// TIA Portal project "M2471_Etiqueteuse" (V18)

(* hardware
DEVICE "Station S7-1200_1"  S7-1200 Station
   slot 0: "Châssis_0"  S7-1200 Rack  Rack  V1.0
   slot 1: "PLC_1"  CPU 1212C DC/DC/DC  6ES7 212-1AE40-0XB0  V4.5
   slot 2: "DI 16/DQ 16x24VDC_1"  6ES7 223-1BL32-0XB0  V2.0
DEVICE "HMI_1"  KTP700 Basic PN
   slot 0: "HMI_1"  KTP700 Basic PN  6AV2 123-2GB03-0AX0  13.0.1.0
   slot 1: "HMI_RT_2"  KTP700 Basic PN  6AV2 123-2GB03-0AX0  13.0.1.0
   slot 5: "HMI_1.IE_CP_1"  PROFINET Interface  13.0.1.0
      slot 1: "Interface PROFINET_1"  PROFINET Interface
         slot 1: "Port_1"  Port
*)

// ===== PLC "PLC_1"  CPU 1212C DC/DC/DC =====

VAR_GLOBAL   // PLC tag table "Table de variables standard"
   "Moteur_Con_Entree" AT %Q8.0 : Bool;
   "Moteur_Con_Etiquetage" AT %Q8.1 : Bool;
   "Moteur_Con_Sortie" AT %Q8.2 : Bool;
   "Moteur_Etiquetage" AT %Q0.7 : Bool;
   "Capteur_Con_Entree" AT %I0.2 : Bool;
   "Capteur_Etiquette" AT %I0.7 : Bool;
   "Capteur_Verin_Tete_Max" AT %I0.4 : Bool;
   "Capteur_Verin_Tete_Min" AT %I0.5 : Bool;
   "Capteur_Verin_Etiquette_Max" AT %I8.0 : Bool;
   "Findecourse_Entree_Petit" AT %I1.6 : Bool;
   "Findecourse_Entree_Grand" AT %I1.7 : Bool;
   "Findecourse_Hauteur_Haut" AT %I0.6 : Bool;
   "Relai_Securite_Arret" AT %I0.0 : Bool;
   "Relai_Secu" AT %Q0.0 : Bool;
   "Moteurpasapas_Haut" AT %M0.0 : Bool;
   "Moteurpasapas_Bas" AT %M0.1 : Bool;
   "Motor_EN" AT %Q0.2 : Bool;
   "Motor_CLK" AT %Q0.4 : Bool;
   "Motor_DIR" AT %Q0.3 : Bool;
   "Entre_Detection_Pot" AT %M0.2 : Bool;
   "Sortie_Detection_Pot" AT %M0.6 : Bool;
   "Butee_Bas_Calibration" AT %I0.1 : Bool;
   "Petit_Pot" AT %M1.0 : Bool;
   "Grand_Pot" AT %M1.1 : Bool;
   "retour_Menu" AT %M0.5 : Bool;
   "System_Byte" AT %MB2 : Byte;
   "FirstScan" AT %M2.0 : Bool;
   "DiagStatusUpdate" AT %M2.1 : Bool;
   "AlwaysTRUE" AT %M2.2 : Bool;
   "AlwaysFALSE" AT %M2.3 : Bool;
   "Clock_Byte" AT %MB3 : Byte;
   "Clock_10Hz" AT %M3.0 : Bool;
   "Clock_5Hz" AT %M3.1 : Bool;
   "Clock_2.5Hz" AT %M3.2 : Bool;
   "Clock_2Hz" AT %M3.3 : Bool;
   "Clock_1.25Hz" AT %M3.4 : Bool;
   "Clock_1Hz" AT %M3.5 : Bool;
   "Clock_0.625Hz" AT %M3.6 : Bool;
   "Clock_0.5Hz" AT %M3.7 : Bool;
   "System_Byte(1)" AT %MB1 : Byte;
   "Moteur_Pwm" AT %Q0.1 : Bool;
   "Controle_Verin" AT %Q8.3 : Bool;
   "Dir_Moteur_15v" AT %Q0.5 : Bool;
   "Detection_Sortie_Bas" AT %M9.2 : Bool;
   "Verin_Etiquette" AT %Q8.4 : Bool;
   "Detection_Entree_Bas" AT %I9.0 : Bool;
   "Detection_Entree_Haut" AT %I9.1 : Bool;
   "Findecourse_Sortie" AT %I9.2 : Bool;
   "Capteur_Position_Pot" AT %I0.3 : Bool;
   "Tag_1" AT %QW1008 : Int;
   "calibration" AT %M1.3 : Bool;
   "stop bourage" AT %M4.0 : Bool;
END_VAR

DATA_BLOCK "Bloc_M2471Etiqueteuse"   // DB1
{ S7_Optimized_Access := 'TRUE' }
VERSION : 0.1
   VAR
      Status_McPower : Bool;
      Hauteur_Haut_Manuel : Bool;
      P_Trig_Reset : Bool;
      Commande_Moteur_Etiquette : Bool;
      Hauteur_Bas_Manuel : Bool;
      Calibrage_Fini : Bool;
      Relai_Securite_Etat : Bool;
      Coordonees_Positionement : Int;
      Moteur_Hauteur_Etiquetage : Bool;
      Moteurpasapas_Sens : Bool;
      Stop_Etat : Bool;
      Moteur_Con_En : Bool;
      Moteur_Con_Et : Bool;
      Moteur_Con_So : Bool;
      Capteur_Entre : Bool;
      capteur_etiquette : Bool;
      Moteur_Etiquette : Bool;
      Capteur_Sortie : Bool;
      Detection_Entre_Petit : Bool;
      Detection_Sortie : Bool;
      Detection_Entre_Grand : Bool;
      Calibration_Home : Bool;
      SR_Home : Bool;
      Ajustement_Hauteur_G_P : Bool;
      Position_Done : Bool;
      Hauteur_Haut_G_P : Bool;
      Hauteur_Bas_G_P : Bool;
      SR_Correction : Bool;
      SR_position : Bool;
      Retour_Menu : Bool;
      Reset : Bool;
      Petit_Pot : Bool;
      Grand_Pot : Bool;
      SR_Position_Done : Bool;
      SR_Correction_Deplacement : Bool;
      Crorrection_Done : Bool;
      Prev_Hauteur_Haut_G_P : Bool;
      Prev_Hauteur_Bas_G_P : Bool;
      Dispense_Etiquette : Bool;
      SR_Etiquette : Bool;
      Etiquetage : Bool;
      P_Trig_Etiquetage : Bool;
      Calibration_set : Bool;
      SR_Home_1 : Bool;
      Sr_etiquetage2 : Bool;
      N_trig_Etiquette : Bool;
      P_trig_Calibration : Bool;
      Reset_Ton_Etiquetage : Bool;
      Controle_Verin_Etiquette : Bool;
      SR_Controle_Verin_Etiquette : Bool;
      Ouverture_Verin_Etiquette : Bool;
      P_trig_Verin_Etiquette : Bool;
      Detection_Petit_Pot : Bool;
      Detection_Grand_Pot : Bool;
      TON_Reset_Controle_Petit : Bool;
      TON_Reset_Controle_Grand : Bool;
      SR_Controle_Petit : Bool;
      SR_Controle_Grand : Bool;
      Sr_Capteur_Pot : Bool;
      P_Trig_Con_Entree : Bool;
      Sr_Capteur_Pot_2 : Bool;
      Sr_Serage_Pot : Bool;
      NTrig_Serage_Pot : Bool;
      SR_CON_Etiquetage : Bool;
      Timer_Con_Etiquetage : Bool;
      Etiquetage_Fini : Bool;
      Verin_Fin : Bool;
      SR_Controle_Verin : Bool;
      SR_Sortie : Bool;
      fin : Bool;
      P_trig_Con_Eti : Bool;
      p_trig_entre : Bool;
      N_trig_etiquetage : Bool;
      controle_Pwm : Bool;
      Machine_Etat : Int;
      Vue_Demarage : Bool;
      Vue_Bourage : Bool;
      Vue_Menu : Bool;
      Vue_Grand : Bool;
      Vue_Petit : Bool;
      Vue_Manuel : Bool;
      Vue_Advance : Bool;
      Bourage : Bool;
      Mise_En_Marche : Bool;
      SR_calibration_Fini : Bool;
      calibrer : Bool;
      Programe : Bool;
      Coordone_Petit_Pot : Int := 100;
      Coordone_Grand_Pot : Int := 160;
      Coordone_Manuel_Pot : Int;
      Confirmation_GP : Bool;
      Confirmation_PP : Bool;
      Pot_Correct : Bool;
      Pot_Incorect : Bool;
      Retour_Demarage : Bool;
      N_Trig_Relai : Bool;
      P_Trig_Reset_calibration : Bool;
      reset_calibration : Bool;
      P_Trig_pot_incorect : Bool;
      SR_Etiquetage_FP : Bool;
      reset_incorect : Bool;
      reset_state : Bool;
      SR_reset : Bool;
      changement_etiquette : Bool;
      nombre_Pot : Int;
      nombre_reset : Bool;
      nombre_limite : Int;
      nombre_Fini : Bool;
      Nombre_sans_limite : Bool;
      p_trigAjustement : Bool;
      p_trig_petit_grand : Bool;
      coordonee_ajustement : Int;
      p_trig_coordone_engage : Bool;
      SR_coordone_engage : Bool;
      p_trig_position_done : Bool;
      p_trig_deplacement : Bool;
      mode_advance : Bool;
      moteur_Grand_advance : Bool;
      moteur_Petit_advance : Bool;
      valeur_Grand_Advance : Int;
      valeur_Petit_Advance : Int;
      coordonne_advance : Int;
      Moteur_advance : Bool;
      Advance_trigger : Bool;
      coordonne_advance_mem : Int;
      valeur_advance_sup_g : Bool;
      valeur_advance_sup_p : Bool;
      p_trig_advance : Bool;
      Manuel_Mode : Bool;
      Manuel_set : Bool;
      Valeur_Manuel : Int;
      Bouton_Manuel_5 : Bool;
      Bouton_Manuel_10 : Bool;
      Bouton_Manuel_25 : Bool;
      Commande_Manuel : Bool;
      Bourage_Done : Bool;
      P_trig_Bourage : Bool;
      bourage_Pneumatique : Bool;
      validation_securite_1 : Bool;
      validation_securite_2 : Bool;
      Verin_Etiquetage : Bool;
      Verin_Etiquette : Bool;
      SR_Bourage_Relai_Secu : Bool;
      Securite_Verin : Bool;
      Home_Reset : Bool;
      p_Trig_Home_Reset : Bool;
      busy_home_Reset : Bool;
      Advance_SR_ajustement : Bool;
      Enable_avdance_Grand : Bool;
      Enable_avdance_Petit : Bool;
      Advance_Etiquetage : Bool;
      SR_Advance : Bool;
      Verin_Etiquetage_advance : Bool;
      Etiquetage_advance : Bool;
      SR_Verin_etiquetage : Bool;
      Bourage_Verin : Bool;
      SR_advance_coordone_done : Bool;
      bourage_verin_etiquette : Bool;
      SR_Grand_Advance : Bool;
      P_trig_Grand_Advance : Bool;
      SR_Petit_Advance : Bool;
      P_trig_Petit_Advance : Bool;
      Grand_Check_Advance : Bool;
      Petit_Check_Advance : Bool;
      Advance_Stop_G : Bool;
      Advance_Stop_P : Bool;
      SR_Controle_P : Bool;
      SR_Controle_G : Bool;
      sr_tapis_eti_fini : Bool;
      reset_Etiquetage : Bool;
      SR_reset_Eti : Bool;
      SR_incorect_tapis_verin : Bool;
      incorect_Reset_P : Bool;
      incorect_Reset_G : Bool;
      sr_con_sortie : Bool;
      Busy_Positionnement : Bool;
      SR_Etiquetage_stop : Bool;
      reset_Absolut_Positionement : Bool;
      error_Positionement : Bool;
      Postionement_reset_error : Bool;
      move_absolut_Busy_Advance : Bool;
      p_trig_advance_Move : Bool;
      p_trig_adv_Etiqu : Bool;
      "SR_advance reset" : Bool;
      SR_Busy_advance_done : Bool;
      advance_check_taille : Int;
      advance_trigger_engage : Bool;
      Sortie_1_etiquette : Bool;
      p_trig_Sortie_1_etiquette : Bool;
      Sr_Advance_fini : Bool;
      advance_move_done : Bool;
      SR_Reset_reset : Bool;
      reset_done : Bool;
      advance_time : Bool;
      advance_time_check : Bool;
      Valeur_manuel_bouton : Bool;
      SR_Manuel_Check : Bool;
      Input_Manuel : Bool;
      P_Trig_Vue_Manuel : Bool;
      reset_Manuel_Check : Bool;
      p_trig_bouton_manuel : Bool;
      insert_Manuel_hauteur : Bool;
      valeur_manuel_check : Int;
      coordoonee_positionement_manuel : Int;
      Etiquetage_comande : Bool;
      reset_sortie_con : Bool;
      SR_reset_con_sortie : Bool;
      p_trig_vue_menu : Bool;
      nouvelle_valeur_manuel : Int;
      comptage_advance_p : Int;
      comptage_advance_g : Int;
      reset_count_p : Bool;
      reset_count_g : Bool;
      bourage_reset : Bool;
      Sr_reset_engage : Bool;
      reset_busy : Bool;
      reset_execute : Bool;
      Sr_reset_done : Bool;
      reset_restart : Bool;
      Home_2_reset : Bool;
      p_trig_home : Bool;
      p_trig_bourage_done : Bool;
      Bourage_Hauteur : Bool;
      p_trig_bourage_hauteur : Bool;
      error_Positionement_Home : Bool;
      error_Positionement_GP : Bool;
      error_Positionement_auto : Bool;
      Fonction_reset : Bool;
      Petit_mem : Bool;
      Grand_mem : Bool;
      checking_taille : Bool;
      automatique_mem : Bool;
      automatique_petit : Bool;
      automatique_grand : Bool;
      set_preset_grand : Bool;
      set_preset_petit : Bool;
   END_VAR
BEGIN
END_DATA_BLOCK

DATA_BLOCK "Initialisation_DB"   // DB2
{ S7_Optimized_Access := 'TRUE' }
VERSION : 0.1
// stored: InstanceOfName Initialisation
"Initialisation"
BEGIN
END_DATA_BLOCK

DATA_BLOCK "En_Marche_DB"   // DB4
{ S7_Optimized_Access := 'TRUE' }
VERSION : 0.1
// stored: InstanceOfName Commande
"Commande"
BEGIN
END_DATA_BLOCK

DATA_BLOCK "HMI_AREA_POINTER"   // DB25
{ S7_Optimized_Access := 'TRUE' }
VERSION : 0.1
   VAR
      tache_API : Array[0..3] of Word;
      NumScreen : Int := 8;
   END_VAR
BEGIN
   tache_API[0] := 51;
   tache_API[2] := 0;
   tache_API[3] := 0;
   // tache_API[1] : Number Screen to display
END_DATA_BLOCK

DATA_BLOCK "Etat_&_Securite_DB"   // DB26
{ S7_Optimized_Access := 'TRUE' }
VERSION : 0.1
// stored: InstanceOfName Etat_&_Securite
"Etat_&_Securite"
BEGIN
END_DATA_BLOCK

DATA_BLOCK "Verin_DB"   // DB28
{ S7_Optimized_Access := 'TRUE' }
VERSION : 0.1
// stored: InstanceOfName Verin
"Verin"
BEGIN
END_DATA_BLOCK

DATA_BLOCK "Moteur_DB"   // DB30
{ S7_Optimized_Access := 'TRUE' }
VERSION : 0.1
// stored: InstanceOfName Moteur
"Moteur"
BEGIN
END_DATA_BLOCK

DATA_BLOCK "Controle_Etiquetage_DB"   // DB31
{ S7_Optimized_Access := 'TRUE' }
VERSION : 0.1
// stored: InstanceOfName Controle_Etiquetage
"Controle_Etiquetage"
BEGIN
END_DATA_BLOCK

DATA_BLOCK "Moteur_DB_1"   // DB35
{ S7_Optimized_Access := 'TRUE' }
VERSION : 0.1
// stored: InstanceOfName Moteur
"Moteur"
BEGIN
END_DATA_BLOCK

DATA_BLOCK "Commande_DB"   // DB37
{ S7_Optimized_Access := 'TRUE' }
VERSION : 0.1
// stored: InstanceOfName Commande
"Commande"
BEGIN
END_DATA_BLOCK

DATA_BLOCK "Commande_DB_1"   // DB38
{ S7_Optimized_Access := 'TRUE' }
VERSION : 0.1
// stored: InstanceOfName Commande
"Commande"
BEGIN
END_DATA_BLOCK

// folder: System blocks/Program resources

DATA_BLOCK "IEC_Timer_0_DB"   // DB5
{ S7_Optimized_Access := 'TRUE' }
AUTHOR : Simatic
FAMILY : IEC
NAME : IEC_TMR
VERSION : 1.0
// stored: InstanceOfName IEC_TIMER
"IEC_TIMER"
BEGIN
END_DATA_BLOCK

DATA_BLOCK "IEC_Counter_0_DB_1"   // DB6
{ S7_Optimized_Access := 'TRUE' }
AUTHOR : Simatic
FAMILY : IEC
NAME : CNTR
VERSION : 1.0
// stored: InstanceOfName IEC_COUNTER
"IEC_COUNTER"
BEGIN
END_DATA_BLOCK

DATA_BLOCK "IEC_Timer_0_DB_2"   // DB7
{ S7_Optimized_Access := 'TRUE' }
AUTHOR : Simatic
FAMILY : IEC
NAME : IEC_TMR
VERSION : 1.0
// stored: InstanceOfName IEC_TIMER
"IEC_TIMER"
BEGIN
END_DATA_BLOCK

DATA_BLOCK "IEC_Timer_0_DB_3"   // DB10
{ S7_Optimized_Access := 'TRUE' }
AUTHOR : Simatic
FAMILY : IEC
NAME : IEC_TMR
VERSION : 1.0
// stored: InstanceOfName IEC_TIMER
"IEC_TIMER"
BEGIN
END_DATA_BLOCK

DATA_BLOCK "IEC_Timer_0_DB_4"   // DB13
{ S7_Optimized_Access := 'TRUE' }
AUTHOR : Simatic
FAMILY : IEC
NAME : IEC_TMR
VERSION : 1.0
// stored: InstanceOfName IEC_TIMER
"IEC_TIMER"
BEGIN
END_DATA_BLOCK

DATA_BLOCK "IEC_Timer_0_DB_5"   // DB15
{ S7_Optimized_Access := 'TRUE' }
AUTHOR : Simatic
FAMILY : IEC
NAME : IEC_TMR
VERSION : 1.0
// stored: InstanceOfName IEC_TIMER
"IEC_TIMER"
BEGIN
END_DATA_BLOCK

DATA_BLOCK "IEC_Counter_0_DB_2"   // DB16
{ S7_Optimized_Access := 'TRUE' }
AUTHOR : Simatic
FAMILY : IEC
NAME : CNTR
VERSION : 1.0
// stored: InstanceOfName IEC_COUNTER
"IEC_COUNTER"
BEGIN
END_DATA_BLOCK

DATA_BLOCK "IEC_Timer_0_DB_7"   // DB17
{ S7_Optimized_Access := 'TRUE' }
AUTHOR : Simatic
FAMILY : IEC
NAME : IEC_TMR
VERSION : 1.0
// stored: InstanceOfName IEC_TIMER
"IEC_TIMER"
BEGIN
END_DATA_BLOCK

DATA_BLOCK "IEC_Timer_0_DB_8"   // DB18
{ S7_Optimized_Access := 'TRUE' }
AUTHOR : Simatic
FAMILY : IEC
NAME : IEC_TMR
VERSION : 1.0
// stored: InstanceOfName IEC_TIMER
"IEC_TIMER"
BEGIN
END_DATA_BLOCK

DATA_BLOCK "IEC_Counter_0_DB"   // DB20
{ S7_Optimized_Access := 'TRUE' }
AUTHOR : Simatic
FAMILY : IEC
NAME : CNTR
VERSION : 1.0
// stored: InstanceOfName IEC_COUNTER
"IEC_COUNTER"
BEGIN
END_DATA_BLOCK

DATA_BLOCK "IEC_Timer_0_DB_9"   // DB27
{ S7_Optimized_Access := 'TRUE' }
AUTHOR : Simatic
FAMILY : IEC
NAME : IEC_TMR
VERSION : 1.0
// stored: InstanceOfName IEC_TIMER
"IEC_TIMER"
BEGIN
END_DATA_BLOCK

DATA_BLOCK "IEC_Timer_0_DB_10"   // DB29
{ S7_Optimized_Access := 'TRUE' }
AUTHOR : Simatic
FAMILY : IEC
NAME : IEC_TMR
VERSION : 1.0
// stored: InstanceOfName IEC_TIMER
"IEC_TIMER"
BEGIN
END_DATA_BLOCK

DATA_BLOCK "IEC_Timer_0_DB_11"   // DB32
{ S7_Optimized_Access := 'TRUE' }
AUTHOR : Simatic
FAMILY : IEC
NAME : IEC_TMR
VERSION : 1.0
// stored: InstanceOfName IEC_TIMER
"IEC_TIMER"
BEGIN
END_DATA_BLOCK

DATA_BLOCK "IEC_Timer_0_DB_12"   // DB34
{ S7_Optimized_Access := 'TRUE' }
AUTHOR : Simatic
FAMILY : IEC
NAME : IEC_TMR
VERSION : 1.0
// stored: InstanceOfName IEC_TIMER
"IEC_TIMER"
BEGIN
END_DATA_BLOCK

DATA_BLOCK "IEC_Timer_0_DB_14"   // DB36
{ S7_Optimized_Access := 'TRUE' }
AUTHOR : Simatic
FAMILY : IEC
NAME : IEC_TMR
VERSION : 1.0
// stored: InstanceOfName IEC_TIMER
"IEC_TIMER"
BEGIN
END_DATA_BLOCK

DATA_BLOCK "IEC_Timer_0_DB_17"   // DB39
{ S7_Optimized_Access := 'TRUE' }
AUTHOR : Simatic
FAMILY : IEC
NAME : IEC_TMR
VERSION : 1.0
// stored: InstanceOfName IEC_TIMER
"IEC_TIMER"
BEGIN
END_DATA_BLOCK

DATA_BLOCK "IEC_Timer_0_DB_18"   // DB40
{ S7_Optimized_Access := 'TRUE' }
AUTHOR : Simatic
FAMILY : IEC
NAME : IEC_TMR
VERSION : 1.0
// stored: InstanceOfName IEC_TIMER
"IEC_TIMER"
BEGIN
END_DATA_BLOCK

DATA_BLOCK "IEC_Timer_0_DB_19"   // DB41
{ S7_Optimized_Access := 'TRUE' }
AUTHOR : Simatic
FAMILY : IEC
NAME : IEC_TMR
VERSION : 1.0
// stored: InstanceOfName IEC_TIMER
"IEC_TIMER"
BEGIN
END_DATA_BLOCK

DATA_BLOCK "IEC_Timer_0_DB_20"   // DB42
{ S7_Optimized_Access := 'TRUE' }
AUTHOR : Simatic
FAMILY : IEC
NAME : IEC_TMR
VERSION : 1.0
// stored: InstanceOfName IEC_TIMER
"IEC_TIMER"
BEGIN
END_DATA_BLOCK

DATA_BLOCK "IEC_Timer_0_DB_21"   // DB45
{ S7_Optimized_Access := 'TRUE' }
AUTHOR : Simatic
FAMILY : IEC
NAME : IEC_TMR
VERSION : 1.0
// stored: InstanceOfName IEC_TIMER
"IEC_TIMER"
BEGIN
END_DATA_BLOCK

DATA_BLOCK "IEC_Timer_0_DB_22"   // DB46
{ S7_Optimized_Access := 'TRUE' }
AUTHOR : Simatic
FAMILY : IEC
NAME : IEC_TMR
VERSION : 1.0
// stored: InstanceOfName IEC_TIMER
"IEC_TIMER"
BEGIN
END_DATA_BLOCK

DATA_BLOCK "IEC_Timer_0_DB_23"   // DB47
{ S7_Optimized_Access := 'TRUE' }
AUTHOR : Simatic
FAMILY : IEC
NAME : IEC_TMR
VERSION : 1.0
// stored: InstanceOfName IEC_TIMER
"IEC_TIMER"
BEGIN
END_DATA_BLOCK

DATA_BLOCK "IEC_Timer_0_DB_24"   // DB48
{ S7_Optimized_Access := 'TRUE' }
AUTHOR : Simatic
FAMILY : IEC
NAME : IEC_TMR
VERSION : 1.0
// stored: InstanceOfName IEC_TIMER
"IEC_TIMER"
BEGIN
END_DATA_BLOCK

// folder: (top level)

DATA_BLOCK "Axe_1"   // DB8, Motion_DB
{ S7_Optimized_Access := 'TRUE' }
AUTHOR : SIMATIC
FAMILY : BasicMC
NAME : TO_PosAx
VERSION : 8.0
// stored: InstanceOfName TO_PositioningAxis
"TO_PositioningAxis"
BEGIN
   // Axis.PositionLimitsMin_AddressCU = %I0.1
   // Axis.PositionLimitsMax_AddressCU = %I0.6
   // Axis.DirectionOutputEnabledCU = TRUE
   // Axis.LengthUnitNormalized.Distance = 1013
   // Axis.HomingReferencePointSwitch_AddressCU = %I0.1
   // Axis.EnableOutput_AddressCU = %Q0.2
   // Axis.OnlinePtoModeCU = 16#0000_0002
   // Axis.SelectedChannel2EnumCU = %Q0.3
   // Axis.SelectedChannel1EnumCU = %Q0.4
   // Pulse.MinDeltaDeltaFrequencyCU = 0.004
   // Pulse.MaxDeltaDeltaFrequencyCU = 1.0E+10
   // Pulse.MinDeltaFrequencyCU = 0.005
   // Pulse.MaxDeltaFrequencyCU = 9.5E+9
   // Pulse.MinFrequencyCU = 1.0
   // Pulse.MaxFrequencyCU = 30000.0
   // Pulse.OutputSourceCU = 16#0000_0000
   // Axis.SelectPTO = 0
END_DATA_BLOCK

FUNCTION_BLOCK "Etat_&_Securite"   // FB1, LAD
{ S7_Optimized_Access := 'TRUE' }
VERSION : 0.1
   VAR_TEMP   // added for the SCL form of the ladder/FBD networks
      _w1 : Bool;
      _w2 : Bool;
   END_VAR
BEGIN

REGION Network 1: Relai de Secrurite
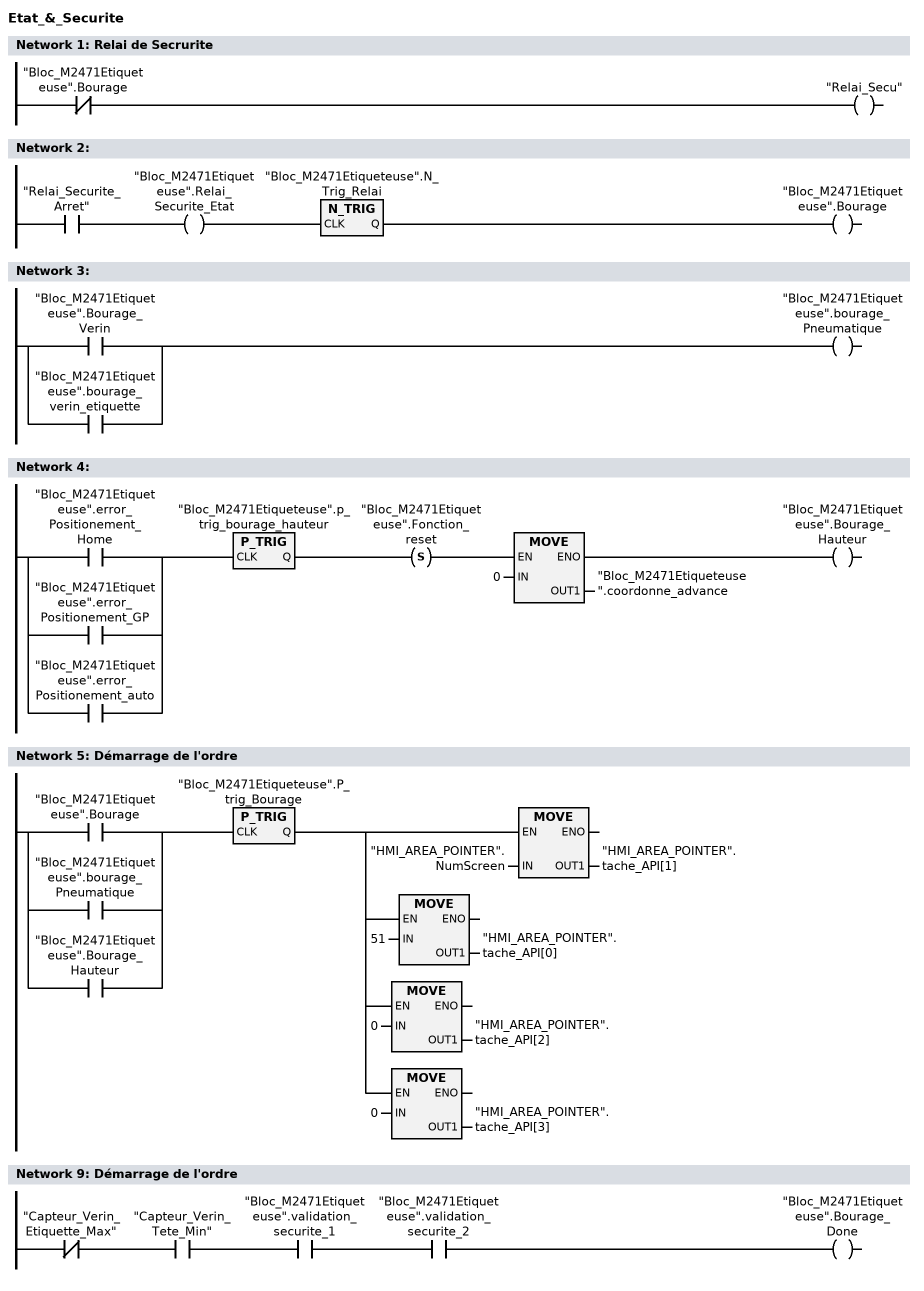
   RUNG wire#powerrail
      I_Contact( "Bloc_M2471Etiqueteuse".Bourage )
      Coil( "Relai_Secu" )
   END_RUNG
   // the same network as SCL:
   "Relai_Secu" := NOT "Bloc_M2471Etiqueteuse".Bourage;
END_REGION

REGION Network 2
   RUNG wire#powerrail
      Contact( "Relai_Securite_Arret" )
      Coil( "Bloc_M2471Etiqueteuse".Relai_Securite_Etat )
      N_Trig( "Bloc_M2471Etiqueteuse".N_Trig_Relai )
      Coil( "Bloc_M2471Etiqueteuse".Bourage )
   END_RUNG
   // the same network as SCL:
   "Bloc_M2471Etiqueteuse".Relai_Securite_Etat := "Relai_Securite_Arret";
   #_w1 := NOT "Relai_Securite_Arret" AND "Bloc_M2471Etiqueteuse".N_Trig_Relai;   // falling edge
   "Bloc_M2471Etiqueteuse".N_Trig_Relai := "Relai_Securite_Arret";
   "Bloc_M2471Etiqueteuse".Bourage := #_w1;
END_REGION

REGION Network 3
   RUNG wire#powerrail
      Contact( "Bloc_M2471Etiqueteuse".Bourage_Verin )
      wire#w1
      Coil( "Bloc_M2471Etiqueteuse".bourage_Pneumatique )
   END_RUNG
   RUNG wire#powerrail
      Contact( "Bloc_M2471Etiqueteuse".bourage_verin_etiquette )
   END_RUNG wire#w1
   // the same network as SCL:
   "Bloc_M2471Etiqueteuse".bourage_Pneumatique := "Bloc_M2471Etiqueteuse".Bourage_Verin OR "Bloc_M2471Etiqueteuse".bourage_verin_etiquette;
END_REGION

REGION Network 4
   RUNG wire#powerrail
      Contact( "Bloc_M2471Etiqueteuse".error_Positionement_Home )
      wire#w1
      P_Trig( "Bloc_M2471Etiqueteuse".p_trig_bourage_hauteur )
      S_Coil( "Bloc_M2471Etiqueteuse".Fonction_reset )
      Move(in := 0, out1 => "Bloc_M2471Etiqueteuse".coordonne_advance)
      Coil( "Bloc_M2471Etiqueteuse".Bourage_Hauteur )
   END_RUNG
   RUNG wire#powerrail
      Contact( "Bloc_M2471Etiqueteuse".error_Positionement_GP )
   END_RUNG wire#w1
   RUNG wire#powerrail
      Contact( "Bloc_M2471Etiqueteuse".error_Positionement_auto )
   END_RUNG wire#w1
   // the same network as SCL:
   #_w1 := "Bloc_M2471Etiqueteuse".error_Positionement_Home OR "Bloc_M2471Etiqueteuse".error_Positionement_GP OR "Bloc_M2471Etiqueteuse".error_Positionement_auto;
   #_w2 := #_w1 AND NOT "Bloc_M2471Etiqueteuse".p_trig_bourage_hauteur;   // rising edge
   "Bloc_M2471Etiqueteuse".p_trig_bourage_hauteur := #_w1;
   IF #_w2 THEN
       "Bloc_M2471Etiqueteuse".Fonction_reset := TRUE;
       "Bloc_M2471Etiqueteuse".coordonne_advance := 0;
   END_IF;
   "Bloc_M2471Etiqueteuse".Bourage_Hauteur := #_w2;
END_REGION

REGION Network 5: Démarrage de l'ordre
   RUNG wire#powerrail
      Contact( "Bloc_M2471Etiqueteuse".Bourage )
      wire#w1
      P_Trig( "Bloc_M2471Etiqueteuse".P_trig_Bourage )
      wire#w2
      Move(in := "HMI_AREA_POINTER".NumScreen, out1 => "HMI_AREA_POINTER".tache_API[1])
   END_RUNG
   RUNG wire#powerrail
      Contact( "Bloc_M2471Etiqueteuse".bourage_Pneumatique )
   END_RUNG wire#w1
   RUNG wire#powerrail
      Contact( "Bloc_M2471Etiqueteuse".Bourage_Hauteur )
   END_RUNG wire#w1
   RUNG wire#w2
      Move(in := 51, out1 => "HMI_AREA_POINTER".tache_API[0])
   END_RUNG
   RUNG wire#w2
      Move(in := 0, out1 => "HMI_AREA_POINTER".tache_API[2])
   END_RUNG
   RUNG wire#w2
      Move(in := 0, out1 => "HMI_AREA_POINTER".tache_API[3])
   END_RUNG
   // the same network as SCL:
   #_w1 := "Bloc_M2471Etiqueteuse".Bourage OR "Bloc_M2471Etiqueteuse".bourage_Pneumatique OR "Bloc_M2471Etiqueteuse".Bourage_Hauteur;
   #_w2 := #_w1 AND NOT "Bloc_M2471Etiqueteuse".P_trig_Bourage;   // rising edge
   "Bloc_M2471Etiqueteuse".P_trig_Bourage := #_w1;
   IF #_w2 THEN
       "HMI_AREA_POINTER".tache_API[1] := "HMI_AREA_POINTER".NumScreen;
       "HMI_AREA_POINTER".tache_API[0] := 51;
       "HMI_AREA_POINTER".tache_API[2] := 0;
       "HMI_AREA_POINTER".tache_API[3] := 0;
   END_IF;
END_REGION

REGION Network 6 (SCL): Machine Etat
   IF "Relai_Securite_Arret" = FALSE OR "Bloc_M2471Etiqueteuse".Bourage OR "Bloc_M2471Etiqueteuse".Bourage_Hauteur OR "Bloc_M2471Etiqueteuse".bourage_Pneumatique OR "Bloc_M2471Etiqueteuse".bourage_reset THEN
       "Bloc_M2471Etiqueteuse".Machine_Etat := 0;

   ELSIF "Bloc_M2471Etiqueteuse".Machine_Etat = 0 AND "Relai_Securite_Arret" = TRUE AND "Bloc_M2471Etiqueteuse".Relai_Securite_Etat = TRUE AND NOT "Bloc_M2471Etiqueteuse".Vue_Bourage =  TRUE THEN
       "Bloc_M2471Etiqueteuse".Machine_Etat := 1;

   ELSIF "Bloc_M2471Etiqueteuse".Machine_Etat = 1 AND "Bloc_M2471Etiqueteuse".calibrer = 1 THEN
      "Bloc_M2471Etiqueteuse".Machine_Etat := 2;

   ELSIF "Bloc_M2471Etiqueteuse".Machine_Etat = 2 AND "Bloc_M2471Etiqueteuse".Programe = 1 THEN
       "Bloc_M2471Etiqueteuse".Machine_Etat := 3;

   ELSIF "Bloc_M2471Etiqueteuse".Machine_Etat = 3 AND "Bloc_M2471Etiqueteuse".Programe = 0 THEN
       "Bloc_M2471Etiqueteuse".Machine_Etat := 2;
   END_IF;
END_REGION

REGION Network 7 (SCL): Etat et Variable
   IF "Bloc_M2471Etiqueteuse".Machine_Etat = 0 THEN
       "Bloc_M2471Etiqueteuse".Calibration_set := 0;
       "Bloc_M2471Etiqueteuse".reset_state := 0;
       "Bloc_M2471Etiqueteuse".Mise_En_Marche := FALSE;

   ELSIF "Bloc_M2471Etiqueteuse".Machine_Etat = 1 THEN
       "Bloc_M2471Etiqueteuse".Fonction_reset :=0;
       "Bloc_M2471Etiqueteuse".Calibration_set := 1;
       "Bloc_M2471Etiqueteuse".reset_state := 0;
       "Bloc_M2471Etiqueteuse".Mise_En_Marche := FALSE;

   ELSIF "Bloc_M2471Etiqueteuse".Machine_Etat = 2 THEN
       "Bloc_M2471Etiqueteuse".Calibration_set := 0;
       "Bloc_M2471Etiqueteuse".reset_state := 0;
       "Bloc_M2471Etiqueteuse".Mise_En_Marche := FALSE;

   ELSIF "Bloc_M2471Etiqueteuse".Machine_Etat = 3 THEN
       "Bloc_M2471Etiqueteuse".reset_state := 1;
       "Bloc_M2471Etiqueteuse".Mise_En_Marche := TRUE;

   END_IF;
END_REGION

REGION Network 8 (SCL): Programmes
   IF "Bloc_M2471Etiqueteuse".Vue_Bourage OR "Bloc_M2471Etiqueteuse".Vue_Demarage = 1 OR "Bloc_M2471Etiqueteuse".Vue_Menu = 1 THEN
       "Bloc_M2471Etiqueteuse".Programe := 0;

   ELSIF "Bloc_M2471Etiqueteuse".Vue_Grand = 1 OR "Bloc_M2471Etiqueteuse".Vue_Petit = 1 OR "Bloc_M2471Etiqueteuse".Vue_Manuel = 1 THEN
       "Bloc_M2471Etiqueteuse".Programe := 1;

   ELSIF "Bloc_M2471Etiqueteuse".Vue_Advance = 1 THEN
       "Bloc_M2471Etiqueteuse".Programe := 1;
       "Bloc_M2471Etiqueteuse".mode_advance := 1;

   END_IF;
END_REGION

REGION Network 9: Démarrage de l'ordre
   RUNG wire#powerrail
      I_Contact( "Capteur_Verin_Etiquette_Max" )
      Contact( "Capteur_Verin_Tete_Min" )
      Contact( "Bloc_M2471Etiqueteuse".validation_securite_1 )
      Contact( "Bloc_M2471Etiqueteuse".validation_securite_2 )
      Coil( "Bloc_M2471Etiqueteuse".Bourage_Done )
   END_RUNG
   // the same network as SCL:
   "Bloc_M2471Etiqueteuse".Bourage_Done := NOT "Capteur_Verin_Etiquette_Max" AND "Capteur_Verin_Tete_Min" AND "Bloc_M2471Etiqueteuse".validation_securite_1 AND "Bloc_M2471Etiqueteuse".validation_securite_2;
END_REGION
END_FUNCTION_BLOCK

FUNCTION_BLOCK "Verin"   // FB2, LAD
{ S7_Optimized_Access := 'TRUE' }
VERSION : 0.1
   VAR_TEMP   // added for the SCL form of the ladder/FBD networks
      _w1 : Bool;
      _w2 : Bool;
      _w3 : Bool;
   END_VAR
BEGIN

REGION Network 1
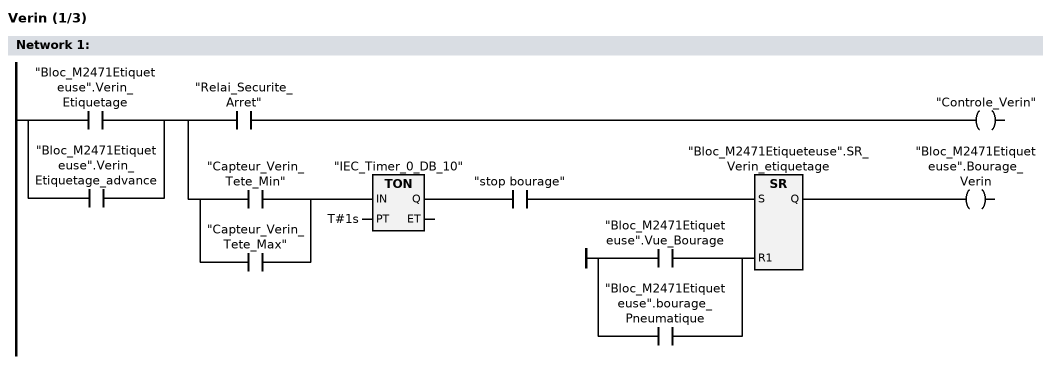
   #_w1 := "Bloc_M2471Etiqueteuse".Verin_Etiquetage OR "Bloc_M2471Etiqueteuse".Verin_Etiquetage_advance;
   "Controle_Verin" := #_w1 AND "Relai_Securite_Arret";
   "IEC_Timer_0_DB_10".TON(IN := #_w1 AND ("Capteur_Verin_Tete_Min" OR "Capteur_Verin_Tete_Max"), PT := T#1s);
   IF "IEC_Timer_0_DB_10".Q AND "stop bourage" THEN
       "Bloc_M2471Etiqueteuse".SR_Verin_etiquetage := TRUE;   // SR flip-flop
   END_IF;
   IF "Bloc_M2471Etiqueteuse".Vue_Bourage OR "Bloc_M2471Etiqueteuse".bourage_Pneumatique THEN
       "Bloc_M2471Etiqueteuse".SR_Verin_etiquetage := FALSE;
   END_IF;
   "Bloc_M2471Etiqueteuse".Bourage_Verin := "Bloc_M2471Etiqueteuse".SR_Verin_etiquetage;
END_REGION

REGION Network 2: commande Pneumatique Verin et tapsi etiquetage
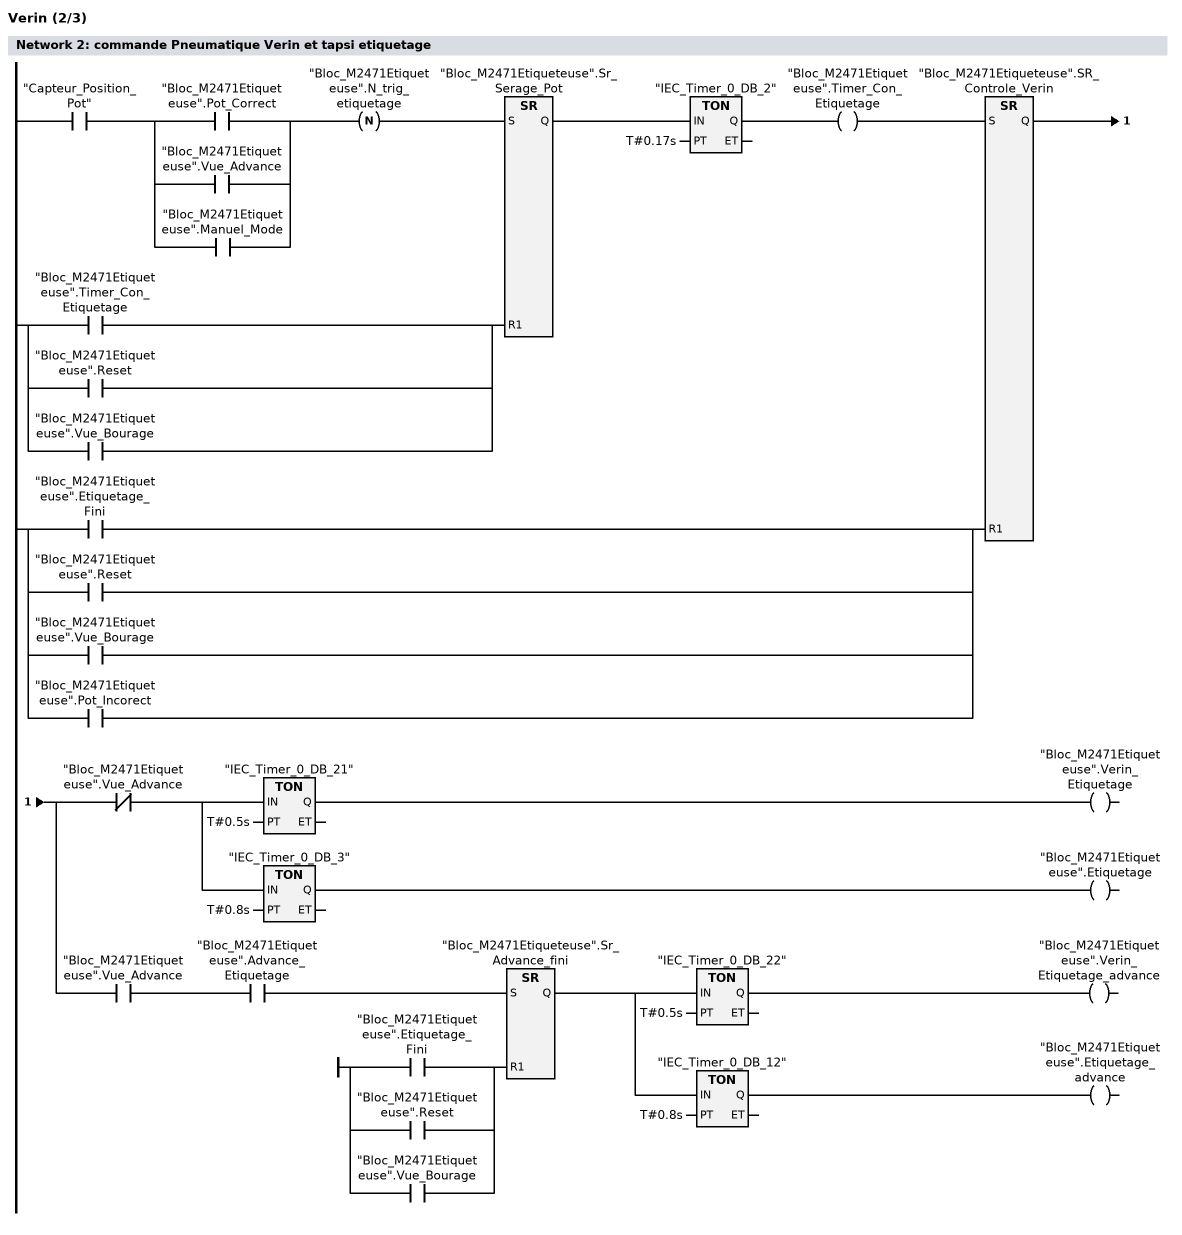
   #_w1 := "Capteur_Position_Pot" AND ("Bloc_M2471Etiqueteuse".Pot_Correct OR "Bloc_M2471Etiqueteuse".Vue_Advance OR "Bloc_M2471Etiqueteuse".Manuel_Mode);
   #_w2 := NOT #_w1 AND "Bloc_M2471Etiqueteuse".N_trig_etiquetage;   // falling edge
   "Bloc_M2471Etiqueteuse".N_trig_etiquetage := #_w1;
   IF #_w2 THEN
       "Bloc_M2471Etiqueteuse".Sr_Serage_Pot := TRUE;   // SR flip-flop
   END_IF;
   IF "Bloc_M2471Etiqueteuse".Timer_Con_Etiquetage OR "Bloc_M2471Etiqueteuse".Reset OR "Bloc_M2471Etiqueteuse".Vue_Bourage THEN
       "Bloc_M2471Etiqueteuse".Sr_Serage_Pot := FALSE;
   END_IF;
   "IEC_Timer_0_DB_2".TON(IN := "Bloc_M2471Etiqueteuse".Sr_Serage_Pot, PT := T#0.17s);
   "Bloc_M2471Etiqueteuse".Timer_Con_Etiquetage := "IEC_Timer_0_DB_2".Q;
   IF "IEC_Timer_0_DB_2".Q THEN
       "Bloc_M2471Etiqueteuse".SR_Controle_Verin := TRUE;   // SR flip-flop
   END_IF;
   IF "Bloc_M2471Etiqueteuse".Etiquetage_Fini OR "Bloc_M2471Etiqueteuse".Reset OR "Bloc_M2471Etiqueteuse".Vue_Bourage OR "Bloc_M2471Etiqueteuse".Pot_Incorect THEN
       "Bloc_M2471Etiqueteuse".SR_Controle_Verin := FALSE;
   END_IF;
   #_w3 := "Bloc_M2471Etiqueteuse".SR_Controle_Verin AND NOT "Bloc_M2471Etiqueteuse".Vue_Advance;
   "IEC_Timer_0_DB_21".TON(IN := #_w3, PT := T#0.5s);
   "Bloc_M2471Etiqueteuse".Verin_Etiquetage := "IEC_Timer_0_DB_21".Q;
   "IEC_Timer_0_DB_3".TON(IN := #_w3, PT := T#0.8s);
   "Bloc_M2471Etiqueteuse".Etiquetage := "IEC_Timer_0_DB_3".Q;
   IF "Bloc_M2471Etiqueteuse".SR_Controle_Verin AND "Bloc_M2471Etiqueteuse".Vue_Advance AND "Bloc_M2471Etiqueteuse".Advance_Etiquetage THEN
       "Bloc_M2471Etiqueteuse".Sr_Advance_fini := TRUE;   // SR flip-flop
   END_IF;
   IF "Bloc_M2471Etiqueteuse".Etiquetage_Fini OR "Bloc_M2471Etiqueteuse".Reset OR "Bloc_M2471Etiqueteuse".Vue_Bourage THEN
       "Bloc_M2471Etiqueteuse".Sr_Advance_fini := FALSE;
   END_IF;
   "IEC_Timer_0_DB_22".TON(IN := "Bloc_M2471Etiqueteuse".Sr_Advance_fini, PT := T#0.5s);
   "Bloc_M2471Etiqueteuse".Verin_Etiquetage_advance := "IEC_Timer_0_DB_22".Q;
   "IEC_Timer_0_DB_12".TON(IN := "Bloc_M2471Etiqueteuse".Sr_Advance_fini, PT := T#0.8s);
   "Bloc_M2471Etiqueteuse".Etiquetage_advance := "IEC_Timer_0_DB_12".Q;
END_REGION

REGION Network 3
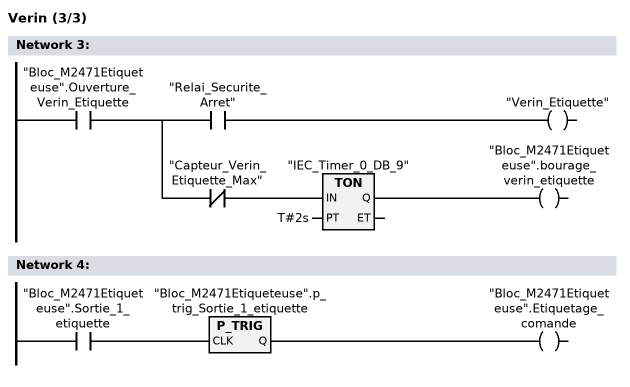
   "Verin_Etiquette" := "Bloc_M2471Etiqueteuse".Ouverture_Verin_Etiquette AND "Relai_Securite_Arret";
   "IEC_Timer_0_DB_9".TON(IN := "Bloc_M2471Etiqueteuse".Ouverture_Verin_Etiquette AND NOT "Capteur_Verin_Etiquette_Max",
                          PT := T#2s);
   "Bloc_M2471Etiqueteuse".bourage_verin_etiquette := "IEC_Timer_0_DB_9".Q;
END_REGION

REGION Network 4
   RUNG wire#powerrail
      Contact( "Bloc_M2471Etiqueteuse".Sortie_1_etiquette )
      P_Trig( "Bloc_M2471Etiqueteuse".p_trig_Sortie_1_etiquette )
      Coil( "Bloc_M2471Etiqueteuse".Etiquetage_comande )
   END_RUNG
   // the same network as SCL:
   #_w1 := "Bloc_M2471Etiqueteuse".Sortie_1_etiquette AND NOT "Bloc_M2471Etiqueteuse".p_trig_Sortie_1_etiquette;   // rising edge
   "Bloc_M2471Etiqueteuse".p_trig_Sortie_1_etiquette := "Bloc_M2471Etiqueteuse".Sortie_1_etiquette;
   "Bloc_M2471Etiqueteuse".Etiquetage_comande := #_w1;
END_REGION
END_FUNCTION_BLOCK

FUNCTION_BLOCK "Commande"   // FB3, LAD
{ S7_Optimized_Access := 'TRUE' }
VERSION : 0.1
   VAR_INPUT
      Valeur_Petit : Int;
      Valeur_Grand : Int;
      Valeur_Ajustement : Int;
   END_VAR
   VAR_TEMP   // added for the SCL form of the ladder/FBD networks
      _w1 : Bool;
   END_VAR
BEGIN

REGION Network 1: Reset
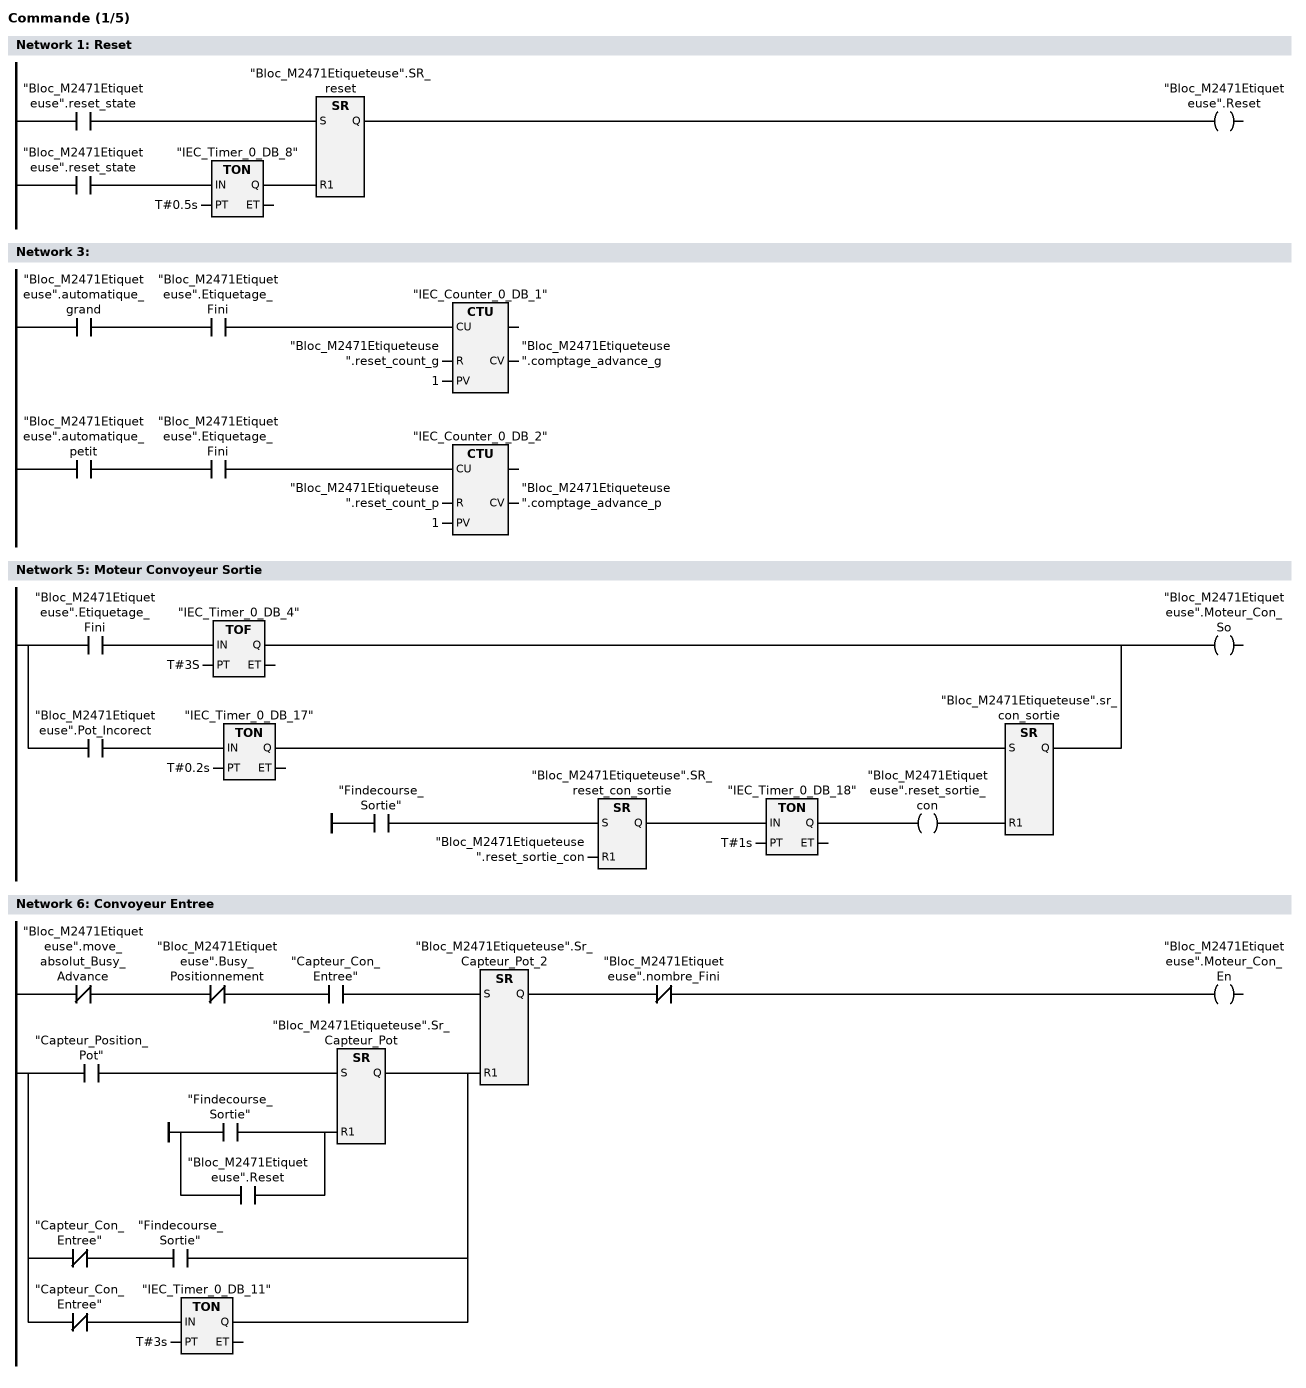
   "IEC_Timer_0_DB_8".TON(IN := "Bloc_M2471Etiqueteuse".reset_state, PT := T#0.5s);
   IF "Bloc_M2471Etiqueteuse".reset_state THEN
       "Bloc_M2471Etiqueteuse".SR_reset := TRUE;   // SR flip-flop
   END_IF;
   IF "IEC_Timer_0_DB_8".Q THEN "Bloc_M2471Etiqueteuse".SR_reset := FALSE; END_IF;
   "Bloc_M2471Etiqueteuse".Reset := "Bloc_M2471Etiqueteuse".SR_reset;
END_REGION

REGION Network 2 (SCL): detection grand ou petit pot ou automatique
   IF "Detection_Entree_Bas" OR "Detection_Entree_Haut" THEN
       "Bloc_M2471Etiqueteuse".checking_taille := 1;
   END_IF;
   IF "Bloc_M2471Etiqueteuse".Vue_Petit THEN
       IF "Detection_Entree_Haut" THEN
           "Bloc_M2471Etiqueteuse".Pot_Incorect := 1;
           "Bloc_M2471Etiqueteuse".Pot_Correct := 0;
           "Bloc_M2471Etiqueteuse".Petit_mem := 1;
       END_IF;
       IF "Bloc_M2471Etiqueteuse".Petit_mem = 0 AND "Bloc_M2471Etiqueteuse".checking_taille  THEN
           "Bloc_M2471Etiqueteuse".Pot_Correct := 1;
           "Bloc_M2471Etiqueteuse".Pot_Incorect := 0;
       END_IF;
   END_IF;

   IF "Bloc_M2471Etiqueteuse".Vue_Grand THEN
       IF "Detection_Entree_Haut" THEN
           "Bloc_M2471Etiqueteuse".Pot_Incorect := 0;
           "Bloc_M2471Etiqueteuse".Pot_Correct := 1;
           "Bloc_M2471Etiqueteuse".Grand_mem := 1;
       END_IF;
       IF "Bloc_M2471Etiqueteuse".Grand_mem = 0 AND "Bloc_M2471Etiqueteuse".checking_taille  THEN
           "Bloc_M2471Etiqueteuse".Pot_Correct := 0;
           "Bloc_M2471Etiqueteuse".Pot_Incorect := 1;
       END_IF;
   END_IF;

   IF "Bloc_M2471Etiqueteuse".Vue_Advance THEN
       IF "Detection_Entree_Haut" AND "Bloc_M2471Etiqueteuse".checking_taille AND "Bloc_M2471Etiqueteuse".automatique_mem = 0 THEN
           "Bloc_M2471Etiqueteuse".moteur_Grand_advance := 1;
           "Bloc_M2471Etiqueteuse".moteur_Petit_advance := 0;
           "Bloc_M2471Etiqueteuse".Advance_Stop_P := 1;
           "Bloc_M2471Etiqueteuse".Advance_Stop_G := 0;
           "Bloc_M2471Etiqueteuse".coordonne_advance := #Valeur_Grand;
           "Bloc_M2471Etiqueteuse".automatique_mem := 1;
           "Bloc_M2471Etiqueteuse".automatique_grand := 1;
           "Bloc_M2471Etiqueteuse".automatique_petit := 0;
       ELSE
           IF "Bloc_M2471Etiqueteuse".checking_taille AND "Bloc_M2471Etiqueteuse".automatique_mem = 0 THEN
               "Bloc_M2471Etiqueteuse".moteur_Grand_advance := 0;
               "Bloc_M2471Etiqueteuse".moteur_Petit_advance := 1;
               "Bloc_M2471Etiqueteuse".Advance_Stop_G := 1;
               "Bloc_M2471Etiqueteuse".Advance_Stop_P := 0;
               "Bloc_M2471Etiqueteuse".coordonne_advance := #Valeur_Petit;
               "Bloc_M2471Etiqueteuse".automatique_grand := 0;
               "Bloc_M2471Etiqueteuse".automatique_petit := 1;
           END_IF;
       END_IF;

   END_IF;
END_REGION

REGION Network 3
   "IEC_Counter_0_DB_1".CTU(CU := "Bloc_M2471Etiqueteuse".automatique_grand AND "Bloc_M2471Etiqueteuse".Etiquetage_Fini,
                           R := "Bloc_M2471Etiqueteuse".reset_count_g,
                           PV := 1,
                           CV => "Bloc_M2471Etiqueteuse".comptage_advance_g);
   "IEC_Counter_0_DB_2".CTU(CU := "Bloc_M2471Etiqueteuse".automatique_petit AND "Bloc_M2471Etiqueteuse".Etiquetage_Fini,
                           R := "Bloc_M2471Etiqueteuse".reset_count_p,
                           PV := 1,
                           CV => "Bloc_M2471Etiqueteuse".comptage_advance_p);
END_REGION

REGION Network 4 (SCL): Pot incorrect RAZBit
   IF "Findecourse_Sortie" = 1 THEN
       "Bloc_M2471Etiqueteuse".Grand_mem := 0;
       "Bloc_M2471Etiqueteuse".Petit_mem := 0;
       "Bloc_M2471Etiqueteuse".automatique_mem := 0;

       "Bloc_M2471Etiqueteuse".checking_taille :=0;
       "Bloc_M2471Etiqueteuse".Pot_Incorect := 0;
       "Bloc_M2471Etiqueteuse".Pot_Correct := 0;

       "Bloc_M2471Etiqueteuse".moteur_Grand_advance := 0;
       "Bloc_M2471Etiqueteuse".moteur_Petit_advance := 0;
       "Bloc_M2471Etiqueteuse".Advance_Stop_G := 1;
       "Bloc_M2471Etiqueteuse".Advance_Stop_P := 1;
       "Bloc_M2471Etiqueteuse".automatique_grand := 0;
       "Bloc_M2471Etiqueteuse".automatique_petit := 0;
   END_IF;
END_REGION

REGION Network 5: Moteur Convoyeur Sortie
   "IEC_Timer_0_DB_4".TOF(IN := "Bloc_M2471Etiqueteuse".Etiquetage_Fini, PT := T#3S);
   "IEC_Timer_0_DB_17".TON(IN := "Bloc_M2471Etiqueteuse".Pot_Incorect, PT := T#0.2s);
   IF "Findecourse_Sortie" THEN
       "Bloc_M2471Etiqueteuse".SR_reset_con_sortie := TRUE;   // SR flip-flop
   END_IF;
   IF "Bloc_M2471Etiqueteuse".reset_sortie_con THEN
       "Bloc_M2471Etiqueteuse".SR_reset_con_sortie := FALSE;
   END_IF;
   "IEC_Timer_0_DB_18".TON(IN := "Bloc_M2471Etiqueteuse".SR_reset_con_sortie, PT := T#1s);
   "Bloc_M2471Etiqueteuse".reset_sortie_con := "IEC_Timer_0_DB_18".Q;
   IF "IEC_Timer_0_DB_17".Q THEN
       "Bloc_M2471Etiqueteuse".sr_con_sortie := TRUE;   // SR flip-flop
   END_IF;
   IF "IEC_Timer_0_DB_18".Q THEN "Bloc_M2471Etiqueteuse".sr_con_sortie := FALSE; END_IF;
   "Bloc_M2471Etiqueteuse".Moteur_Con_So := "IEC_Timer_0_DB_4".Q OR "Bloc_M2471Etiqueteuse".sr_con_sortie;
END_REGION

REGION Network 6: Convoyeur Entree
   IF "Capteur_Position_Pot" THEN
       "Bloc_M2471Etiqueteuse".Sr_Capteur_Pot := TRUE;   // SR flip-flop
   END_IF;
   IF "Findecourse_Sortie" OR "Bloc_M2471Etiqueteuse".Reset THEN
       "Bloc_M2471Etiqueteuse".Sr_Capteur_Pot := FALSE;
   END_IF;
   "IEC_Timer_0_DB_11".TON(IN := NOT "Capteur_Con_Entree", PT := T#3s);
   IF NOT "Bloc_M2471Etiqueteuse".move_absolut_Busy_Advance AND NOT "Bloc_M2471Etiqueteuse".Busy_Positionnement AND "Capteur_Con_Entree" THEN
       "Bloc_M2471Etiqueteuse".Sr_Capteur_Pot_2 := TRUE;   // SR flip-flop
   END_IF;
   IF "Bloc_M2471Etiqueteuse".Sr_Capteur_Pot OR (NOT "Capteur_Con_Entree" AND "Findecourse_Sortie") OR "IEC_Timer_0_DB_11".Q THEN
       "Bloc_M2471Etiqueteuse".Sr_Capteur_Pot_2 := FALSE;
   END_IF;
   "Bloc_M2471Etiqueteuse".Moteur_Con_En := "Bloc_M2471Etiqueteuse".Sr_Capteur_Pot_2 AND NOT "Bloc_M2471Etiqueteuse".nombre_Fini;
END_REGION

REGION Network 7: Convoyeur Etiquetage et timer
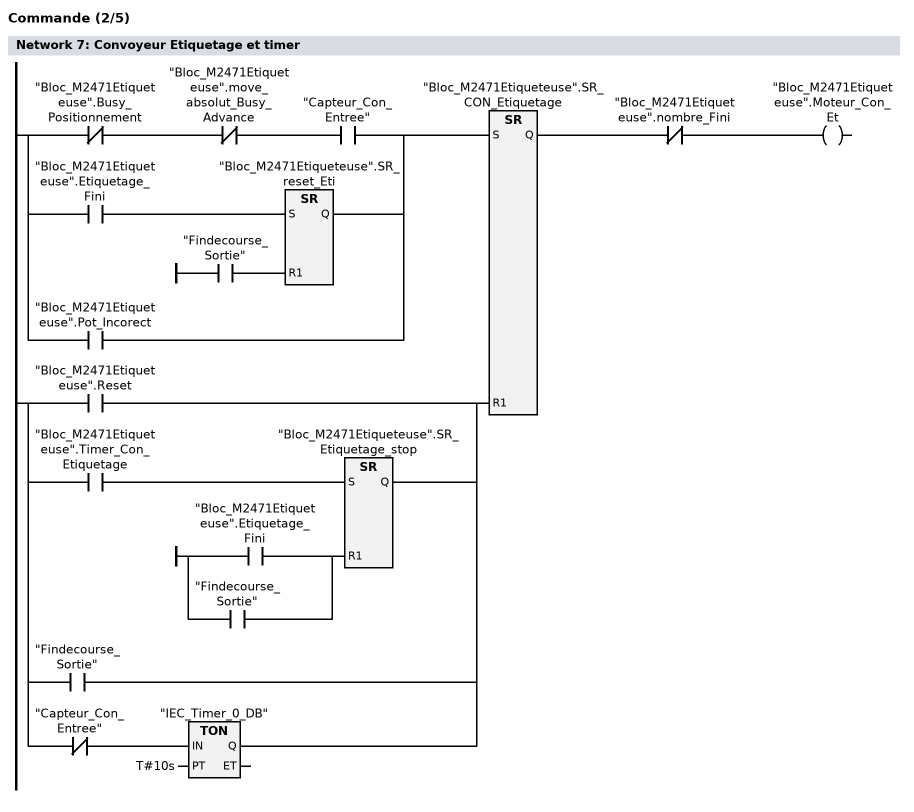
   IF "Bloc_M2471Etiqueteuse".Etiquetage_Fini THEN
       "Bloc_M2471Etiqueteuse".SR_reset_Eti := TRUE;   // SR flip-flop
   END_IF;
   IF "Findecourse_Sortie" THEN "Bloc_M2471Etiqueteuse".SR_reset_Eti := FALSE; END_IF;
   IF "Bloc_M2471Etiqueteuse".Timer_Con_Etiquetage THEN
       "Bloc_M2471Etiqueteuse".SR_Etiquetage_stop := TRUE;   // SR flip-flop
   END_IF;
   IF "Bloc_M2471Etiqueteuse".Etiquetage_Fini OR "Findecourse_Sortie" THEN
       "Bloc_M2471Etiqueteuse".SR_Etiquetage_stop := FALSE;
   END_IF;
   "IEC_Timer_0_DB".TON(IN := NOT "Capteur_Con_Entree", PT := T#10s);
   IF (NOT "Bloc_M2471Etiqueteuse".Busy_Positionnement AND NOT "Bloc_M2471Etiqueteuse".move_absolut_Busy_Advance AND "Capteur_Con_Entree") OR "Bloc_M2471Etiqueteuse".SR_reset_Eti OR "Bloc_M2471Etiqueteuse".Pot_Incorect THEN
       "Bloc_M2471Etiqueteuse".SR_CON_Etiquetage := TRUE;   // SR flip-flop
   END_IF;
   IF "Bloc_M2471Etiqueteuse".Reset OR "Bloc_M2471Etiqueteuse".SR_Etiquetage_stop OR "Findecourse_Sortie" OR "IEC_Timer_0_DB".Q THEN
       "Bloc_M2471Etiqueteuse".SR_CON_Etiquetage := FALSE;
   END_IF;
   "Bloc_M2471Etiqueteuse".Moteur_Con_Et := "Bloc_M2471Etiqueteuse".SR_CON_Etiquetage AND NOT "Bloc_M2471Etiqueteuse".nombre_Fini;
END_REGION

REGION Network 8 (SCL): Controle Hauteur Manuel
   IF  "Bloc_M2471Etiqueteuse".Hauteur_Haut_Manuel = TRUE THEN
       "Bloc_M2471Etiqueteuse".Moteur_Hauteur_Etiquetage:= TRUE;
   ELSIF  "Bloc_M2471Etiqueteuse".Hauteur_Bas_Manuel = TRUE THEN
       "Bloc_M2471Etiqueteuse".Moteur_Hauteur_Etiquetage := TRUE;
   ELSE
       "Bloc_M2471Etiqueteuse".Moteur_Hauteur_Etiquetage := FALSE;
   END_IF;
END_REGION

REGION Network 9 (SCL): Coordonnes Grand ou Petit programe
   "R_TRIG_DB_3"(CLK:="Bloc_M2471Etiqueteuse".Petit_Pot);
   "R_TRIG_DB_4"(CLK:="Bloc_M2471Etiqueteuse".Grand_Pot);
   IF "R_TRIG_DB_3".Q THEN
       "Bloc_M2471Etiqueteuse".Coordonees_Positionement := #Valeur_Petit;
   ELSIF "R_TRIG_DB_4".Q THEN
       "Bloc_M2471Etiqueteuse".Coordonees_Positionement := #Valeur_Grand;
   END_IF;
END_REGION

REGION Network 10: MC_moveabsolut pour Grand ou Petit et manuel
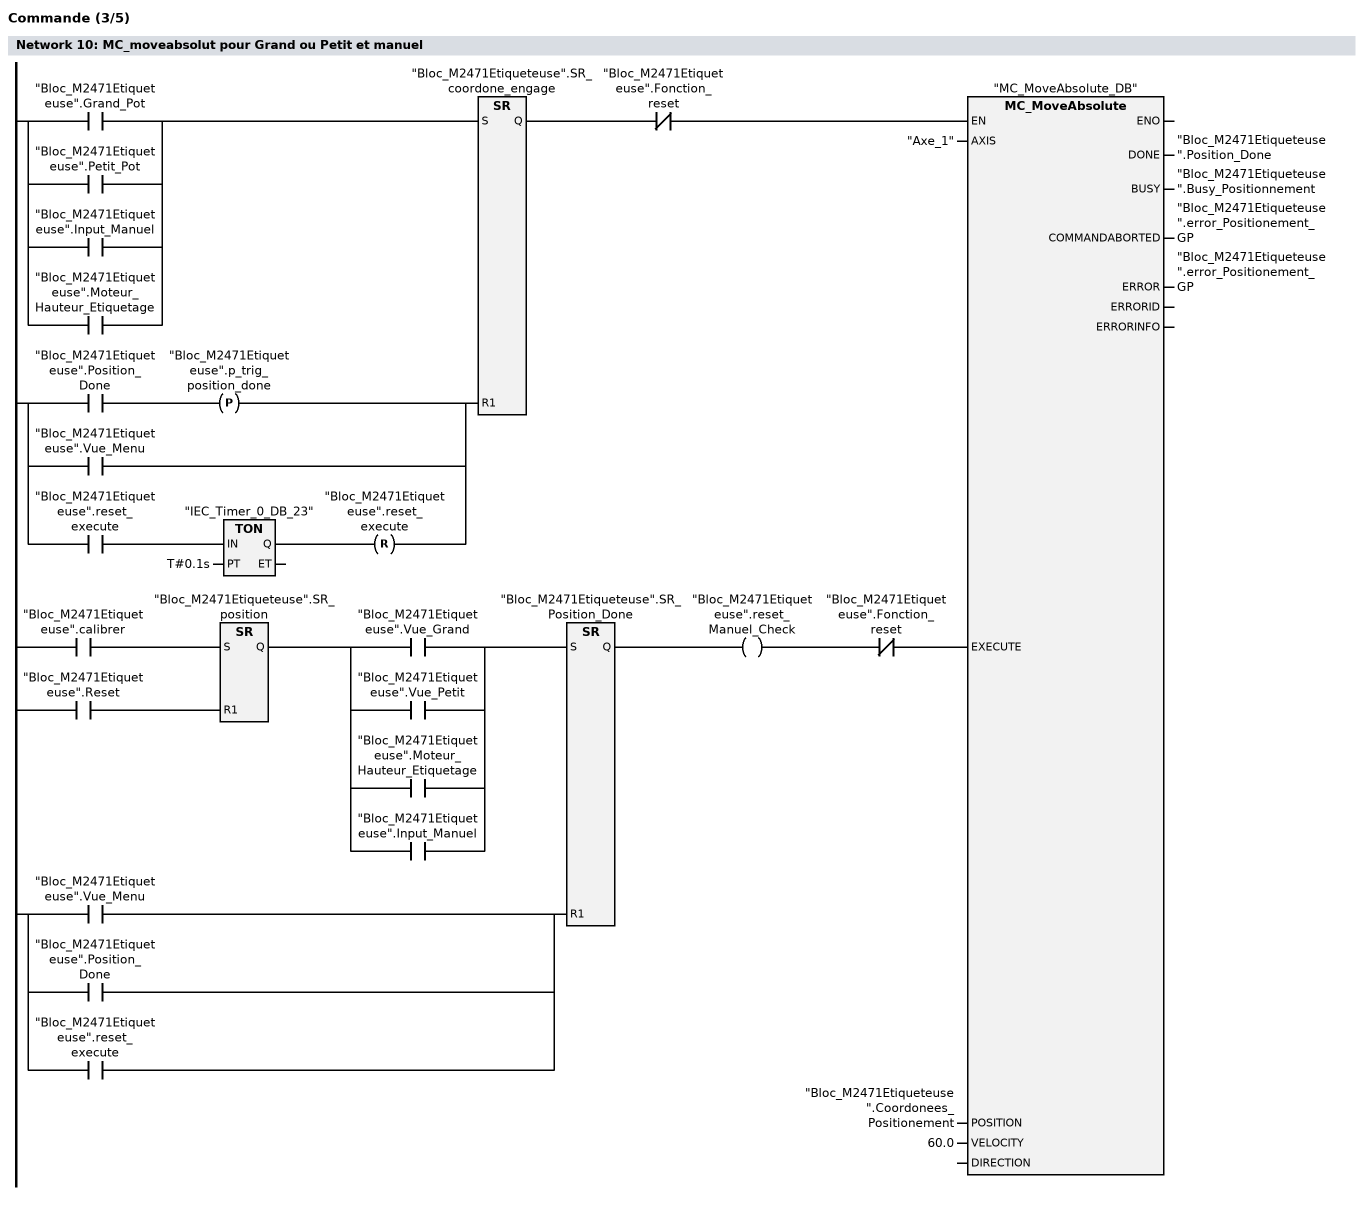
   #_w1 := "Bloc_M2471Etiqueteuse".Position_Done AND NOT "Bloc_M2471Etiqueteuse".p_trig_position_done;   // rising edge
   "Bloc_M2471Etiqueteuse".p_trig_position_done := "Bloc_M2471Etiqueteuse".Position_Done;
   "IEC_Timer_0_DB_23".TON(IN := "Bloc_M2471Etiqueteuse".reset_execute, PT := T#0.1s);
   IF "IEC_Timer_0_DB_23".Q THEN "Bloc_M2471Etiqueteuse".reset_execute := FALSE; END_IF;
   IF "Bloc_M2471Etiqueteuse".Grand_Pot OR "Bloc_M2471Etiqueteuse".Petit_Pot OR "Bloc_M2471Etiqueteuse".Input_Manuel OR "Bloc_M2471Etiqueteuse".Moteur_Hauteur_Etiquetage THEN
       "Bloc_M2471Etiqueteuse".SR_coordone_engage := TRUE;   // SR flip-flop
   END_IF;
   IF #_w1 OR "Bloc_M2471Etiqueteuse".Vue_Menu OR "IEC_Timer_0_DB_23".Q THEN
       "Bloc_M2471Etiqueteuse".SR_coordone_engage := FALSE;
   END_IF;
   IF "Bloc_M2471Etiqueteuse".calibrer THEN
       "Bloc_M2471Etiqueteuse".SR_position := TRUE;   // SR flip-flop
   END_IF;
   IF "Bloc_M2471Etiqueteuse".Reset THEN "Bloc_M2471Etiqueteuse".SR_position := FALSE; END_IF;
   IF "Bloc_M2471Etiqueteuse".SR_position AND ("Bloc_M2471Etiqueteuse".Vue_Grand OR "Bloc_M2471Etiqueteuse".Vue_Petit OR "Bloc_M2471Etiqueteuse".Moteur_Hauteur_Etiquetage OR "Bloc_M2471Etiqueteuse".Input_Manuel) THEN
       "Bloc_M2471Etiqueteuse".SR_Position_Done := TRUE;   // SR flip-flop
   END_IF;
   IF "Bloc_M2471Etiqueteuse".Vue_Menu OR "Bloc_M2471Etiqueteuse".Position_Done OR "Bloc_M2471Etiqueteuse".reset_execute THEN
       "Bloc_M2471Etiqueteuse".SR_Position_Done := FALSE;
   END_IF;
   "Bloc_M2471Etiqueteuse".reset_Manuel_Check := "Bloc_M2471Etiqueteuse".SR_Position_Done;
   IF "Bloc_M2471Etiqueteuse".SR_coordone_engage AND NOT "Bloc_M2471Etiqueteuse".Fonction_reset THEN
       "MC_MoveAbsolute_DB"(Axis := "Axe_1",   // MC_MoveAbsolute
                            Execute := "Bloc_M2471Etiqueteuse".SR_Position_Done AND NOT "Bloc_M2471Etiqueteuse".Fonction_reset,
                            Position := "Bloc_M2471Etiqueteuse".Coordonees_Positionement,
                            Velocity := 60.0,
                            Done => "Bloc_M2471Etiqueteuse".Position_Done,
                            Busy => "Bloc_M2471Etiqueteuse".Busy_Positionnement,
                            CommandAborted => "Bloc_M2471Etiqueteuse".error_Positionement_GP,
                            Error => "Bloc_M2471Etiqueteuse".error_Positionement_GP);
   END_IF;
END_REGION

REGION Network 11: Manuel coordonee
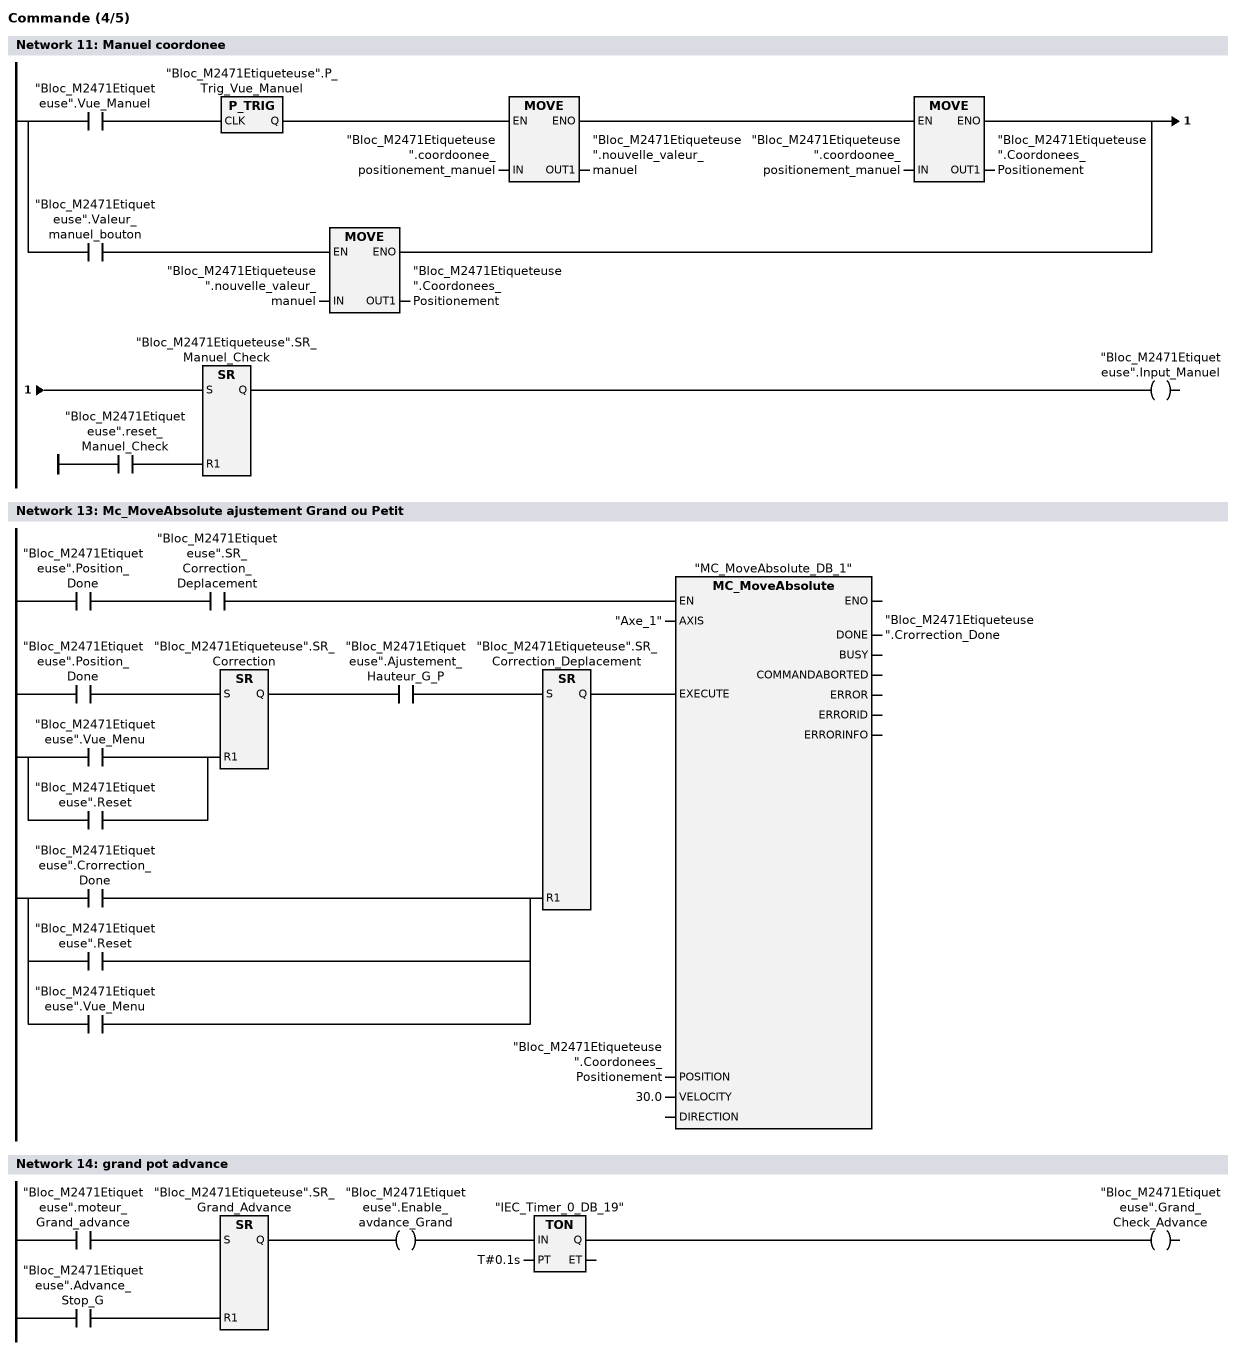
   RUNG wire#powerrail
      Contact( "Bloc_M2471Etiqueteuse".Vue_Manuel )
      P_Trig( "Bloc_M2471Etiqueteuse".P_Trig_Vue_Manuel )
      Move(in := "Bloc_M2471Etiqueteuse".coordoonee_positionement_manuel, out1 => "Bloc_M2471Etiqueteuse".nouvelle_valeur_manuel)
      Move(in := "Bloc_M2471Etiqueteuse".coordoonee_positionement_manuel, out1 => "Bloc_M2471Etiqueteuse".Coordonees_Positionement)
      wire#w1
      S_SR(operand := "Bloc_M2471Etiqueteuse".SR_Manuel_Check, r1 := wire#w2)
      Coil( "Bloc_M2471Etiqueteuse".Input_Manuel )
   END_RUNG
   RUNG wire#powerrail
      Contact( "Bloc_M2471Etiqueteuse".Valeur_manuel_bouton )
      Move(in := "Bloc_M2471Etiqueteuse".nouvelle_valeur_manuel, out1 => "Bloc_M2471Etiqueteuse".Coordonees_Positionement)
   END_RUNG wire#w1
   RUNG wire#powerrail
      Contact( "Bloc_M2471Etiqueteuse".reset_Manuel_Check )
   END_RUNG wire#w2
   // the same network as SCL:
   #_w1 := "Bloc_M2471Etiqueteuse".Vue_Manuel AND NOT "Bloc_M2471Etiqueteuse".P_Trig_Vue_Manuel;   // rising edge
   "Bloc_M2471Etiqueteuse".P_Trig_Vue_Manuel := "Bloc_M2471Etiqueteuse".Vue_Manuel;
   IF #_w1 THEN
       "Bloc_M2471Etiqueteuse".nouvelle_valeur_manuel := "Bloc_M2471Etiqueteuse".coordoonee_positionement_manuel;
       "Bloc_M2471Etiqueteuse".Coordonees_Positionement := "Bloc_M2471Etiqueteuse".coordoonee_positionement_manuel;
   END_IF;
   IF "Bloc_M2471Etiqueteuse".Valeur_manuel_bouton THEN
       "Bloc_M2471Etiqueteuse".Coordonees_Positionement := "Bloc_M2471Etiqueteuse".nouvelle_valeur_manuel;
   END_IF;
   IF #_w1 OR "Bloc_M2471Etiqueteuse".Valeur_manuel_bouton THEN
       "Bloc_M2471Etiqueteuse".SR_Manuel_Check := TRUE;   // SR flip-flop
   END_IF;
   IF "Bloc_M2471Etiqueteuse".reset_Manuel_Check THEN
       "Bloc_M2471Etiqueteuse".SR_Manuel_Check := FALSE;
   END_IF;
   "Bloc_M2471Etiqueteuse".Input_Manuel := "Bloc_M2471Etiqueteuse".SR_Manuel_Check;
END_REGION

REGION Network 12 (SCL): detection fleche haut ou bas
   "R_TRIG_DB_1"(CLK := "Bloc_M2471Etiqueteuse".Hauteur_Haut_Manuel OR "Bloc_M2471Etiqueteuse".Hauteur_Haut_G_P);
   "R_TRIG_DB_2"(CLK:="Bloc_M2471Etiqueteuse".Hauteur_Bas_Manuel OR "Bloc_M2471Etiqueteuse".Hauteur_Bas_G_P);

   IF "R_TRIG_DB_1".Q THEN
       IF NOT "Bloc_M2471Etiqueteuse".Vue_Manuel THEN
           "Bloc_M2471Etiqueteuse".Coordonees_Positionement := "Bloc_M2471Etiqueteuse".Coordonees_Positionement + #Valeur_Ajustement;
       ELSE
           "Bloc_M2471Etiqueteuse".Coordonees_Positionement := "Bloc_M2471Etiqueteuse".Coordonees_Positionement + "Bloc_M2471Etiqueteuse".Valeur_Manuel ;
           "Bloc_M2471Etiqueteuse".insert_Manuel_hauteur := 1;
       END_IF;
       //
   ELSIF "R_TRIG_DB_2".Q THEN
       IF NOT "Bloc_M2471Etiqueteuse".Vue_Manuel THEN
           "Bloc_M2471Etiqueteuse".Coordonees_Positionement := "Bloc_M2471Etiqueteuse".Coordonees_Positionement - #Valeur_Ajustement;
       ELSE
           "Bloc_M2471Etiqueteuse".Coordonees_Positionement := "Bloc_M2471Etiqueteuse".Coordonees_Positionement - "Bloc_M2471Etiqueteuse".Valeur_Manuel;
           "Bloc_M2471Etiqueteuse".insert_Manuel_hauteur := 1;
       END_IF;
   END_IF;
   //
   //
END_REGION

REGION Network 13: Mc_MoveAbsolute ajustement Grand ou Petit
   IF "Bloc_M2471Etiqueteuse".Position_Done THEN
       "Bloc_M2471Etiqueteuse".SR_Correction := TRUE;   // SR flip-flop
   END_IF;
   IF "Bloc_M2471Etiqueteuse".Vue_Menu OR "Bloc_M2471Etiqueteuse".Reset THEN
       "Bloc_M2471Etiqueteuse".SR_Correction := FALSE;
   END_IF;
   #_w1 := "Bloc_M2471Etiqueteuse".Position_Done AND "Bloc_M2471Etiqueteuse".SR_Correction_Deplacement;
   IF "Bloc_M2471Etiqueteuse".SR_Correction AND "Bloc_M2471Etiqueteuse".Ajustement_Hauteur_G_P THEN
       "Bloc_M2471Etiqueteuse".SR_Correction_Deplacement := TRUE;   // SR flip-flop
   END_IF;
   IF "Bloc_M2471Etiqueteuse".Crorrection_Done OR "Bloc_M2471Etiqueteuse".Reset OR "Bloc_M2471Etiqueteuse".Vue_Menu THEN
       "Bloc_M2471Etiqueteuse".SR_Correction_Deplacement := FALSE;
   END_IF;
   IF #_w1 THEN
       "MC_MoveAbsolute_DB_1"(Axis := "Axe_1",   // MC_MoveAbsolute
                              Execute := "Bloc_M2471Etiqueteuse".SR_Correction_Deplacement,
                              Position := "Bloc_M2471Etiqueteuse".Coordonees_Positionement,
                              Velocity := 30.0,
                              Done => "Bloc_M2471Etiqueteuse".Crorrection_Done);
   END_IF;
END_REGION

REGION Network 14: grand pot advance
   IF "Bloc_M2471Etiqueteuse".moteur_Grand_advance THEN
       "Bloc_M2471Etiqueteuse".SR_Grand_Advance := TRUE;   // SR flip-flop
   END_IF;
   IF "Bloc_M2471Etiqueteuse".Advance_Stop_G THEN "Bloc_M2471Etiqueteuse".SR_Grand_Advance := FALSE; END_IF;
   "Bloc_M2471Etiqueteuse".Enable_avdance_Grand := "Bloc_M2471Etiqueteuse".SR_Grand_Advance;
   "IEC_Timer_0_DB_19".TON(IN := "Bloc_M2471Etiqueteuse".SR_Grand_Advance, PT := T#0.1s);
   "Bloc_M2471Etiqueteuse".Grand_Check_Advance := "IEC_Timer_0_DB_19".Q;
END_REGION

REGION Network 15: petit pot advance
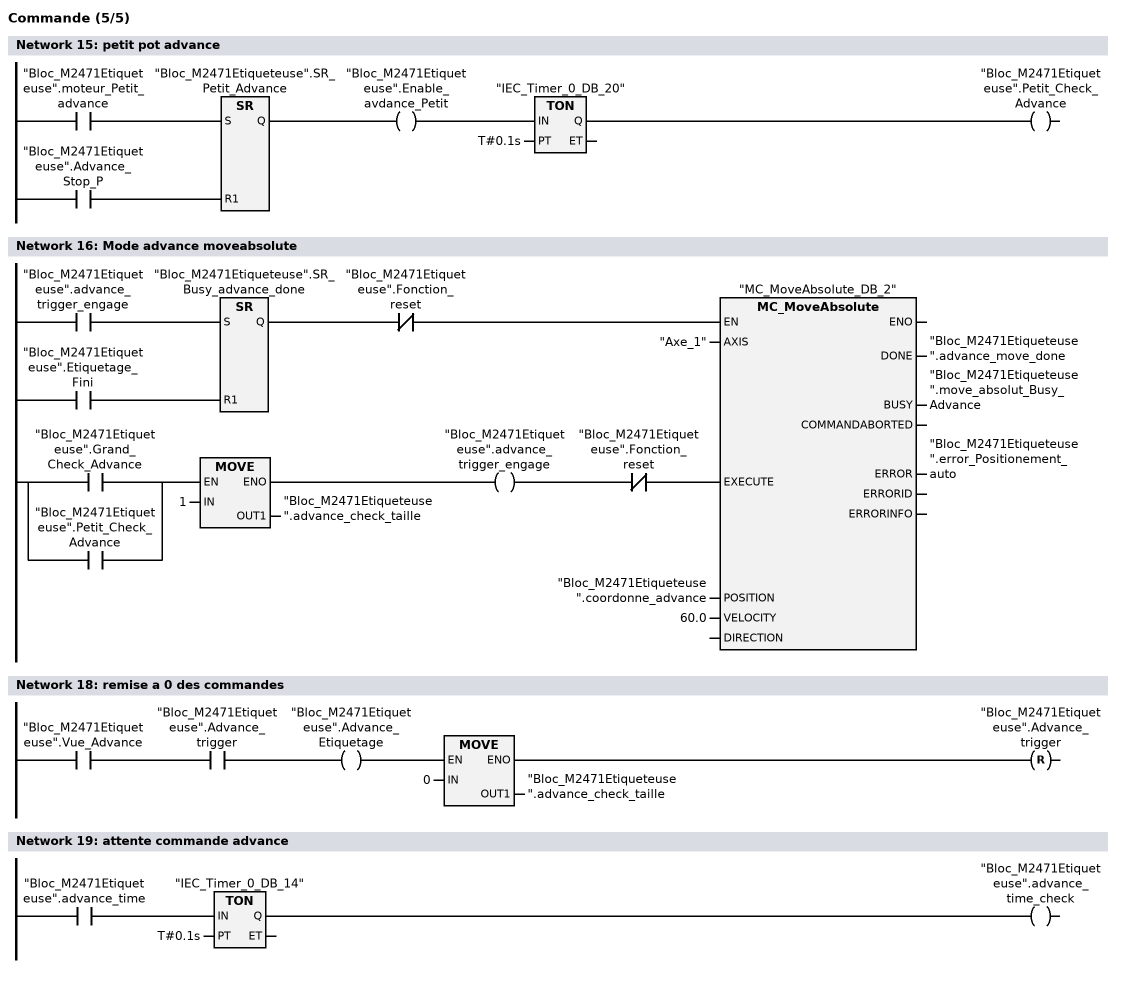
   IF "Bloc_M2471Etiqueteuse".moteur_Petit_advance THEN
       "Bloc_M2471Etiqueteuse".SR_Petit_Advance := TRUE;   // SR flip-flop
   END_IF;
   IF "Bloc_M2471Etiqueteuse".Advance_Stop_P THEN "Bloc_M2471Etiqueteuse".SR_Petit_Advance := FALSE; END_IF;
   "Bloc_M2471Etiqueteuse".Enable_avdance_Petit := "Bloc_M2471Etiqueteuse".SR_Petit_Advance;
   "IEC_Timer_0_DB_20".TON(IN := "Bloc_M2471Etiqueteuse".SR_Petit_Advance, PT := T#0.1s);
   "Bloc_M2471Etiqueteuse".Petit_Check_Advance := "IEC_Timer_0_DB_20".Q;
END_REGION

REGION Network 16: Mode advance moveabsolute
   IF "Bloc_M2471Etiqueteuse".advance_trigger_engage THEN
       "Bloc_M2471Etiqueteuse".SR_Busy_advance_done := TRUE;   // SR flip-flop
   END_IF;
   IF "Bloc_M2471Etiqueteuse".Etiquetage_Fini THEN
       "Bloc_M2471Etiqueteuse".SR_Busy_advance_done := FALSE;
   END_IF;
   #_w1 := "Bloc_M2471Etiqueteuse".Grand_Check_Advance OR "Bloc_M2471Etiqueteuse".Petit_Check_Advance;
   IF #_w1 THEN "Bloc_M2471Etiqueteuse".advance_check_taille := 1; END_IF;
   "Bloc_M2471Etiqueteuse".advance_trigger_engage := #_w1;
   IF "Bloc_M2471Etiqueteuse".SR_Busy_advance_done AND NOT "Bloc_M2471Etiqueteuse".Fonction_reset THEN
       "MC_MoveAbsolute_DB_2"(Axis := "Axe_1",   // MC_MoveAbsolute
                              Execute := #_w1 AND NOT "Bloc_M2471Etiqueteuse".Fonction_reset,
                              Position := "Bloc_M2471Etiqueteuse".coordonne_advance,
                              Velocity := 60.0,
                              Done => "Bloc_M2471Etiqueteuse".advance_move_done,
                              Busy => "Bloc_M2471Etiqueteuse".move_absolut_Busy_Advance,
                              Error => "Bloc_M2471Etiqueteuse".error_Positionement_auto);
   END_IF;
END_REGION

REGION Network 17 (SCL): Detection de difference d'hauteur
   IF "Bloc_M2471Etiqueteuse".advance_check_taille = 1 THEN
       IF "Bloc_M2471Etiqueteuse".coordonne_advance <> "Bloc_M2471Etiqueteuse".coordonne_advance_mem THEN
           "Bloc_M2471Etiqueteuse".advance_time := 1;
           IF "Bloc_M2471Etiqueteuse".move_absolut_Busy_Advance = 1 AND "Bloc_M2471Etiqueteuse".advance_move_done =0 THEN
               "Bloc_M2471Etiqueteuse".Advance_trigger := 0;
           ELSIF "Bloc_M2471Etiqueteuse".advance_time_check = 1 THEN
               "Bloc_M2471Etiqueteuse".coordonne_advance_mem := "Bloc_M2471Etiqueteuse".coordonne_advance;
               "Bloc_M2471Etiqueteuse".Advance_trigger := 1;
               "Bloc_M2471Etiqueteuse".advance_time := 0;
           END_IF;
       ELSE
           "Bloc_M2471Etiqueteuse".coordonne_advance_mem := "Bloc_M2471Etiqueteuse".coordonne_advance;
           "Bloc_M2471Etiqueteuse".Advance_trigger := 1;
       END_IF;
   ELSE
       ;
   END_IF;
END_REGION

REGION Network 18: remise a 0 des commandes
   RUNG wire#powerrail
      Contact( "Bloc_M2471Etiqueteuse".Vue_Advance )
      Contact( "Bloc_M2471Etiqueteuse".Advance_trigger )
      Coil( "Bloc_M2471Etiqueteuse".Advance_Etiquetage )
      Move(in := 0, out1 => "Bloc_M2471Etiqueteuse".advance_check_taille)
      R_Coil( "Bloc_M2471Etiqueteuse".Advance_trigger )
   END_RUNG
   // the same network as SCL:
   "Bloc_M2471Etiqueteuse".Advance_Etiquetage := "Bloc_M2471Etiqueteuse".Vue_Advance AND "Bloc_M2471Etiqueteuse".Advance_trigger;
   IF "Bloc_M2471Etiqueteuse".Advance_Etiquetage THEN
       "Bloc_M2471Etiqueteuse".advance_check_taille := 0;
       "Bloc_M2471Etiqueteuse".Advance_trigger := FALSE;
   END_IF;
END_REGION

REGION Network 19: attente commande advance
   "IEC_Timer_0_DB_14".TON(IN := "Bloc_M2471Etiqueteuse".advance_time, PT := T#0.1s);
   "Bloc_M2471Etiqueteuse".advance_time_check := "IEC_Timer_0_DB_14".Q;
END_REGION
END_FUNCTION_BLOCK

FUNCTION_BLOCK "Moteur"   // FB4, LAD
{ S7_Optimized_Access := 'TRUE' }
VERSION : 0.1
BEGIN

REGION Network 1: Controle_PWM
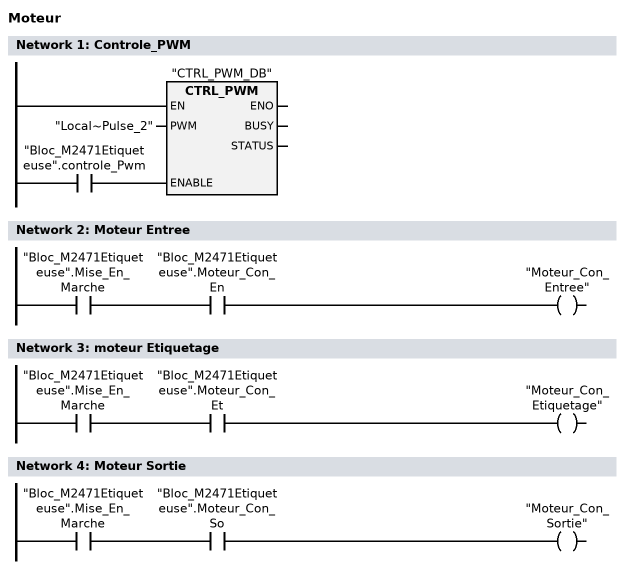
   "CTRL_PWM_DB"(PWM := "Local~Pulse_2", ENABLE := "Bloc_M2471Etiqueteuse".controle_Pwm);   // CTRL_PWM
END_REGION

REGION Network 2: Moteur Entree
   RUNG wire#powerrail
      Contact( "Bloc_M2471Etiqueteuse".Mise_En_Marche )
      Contact( "Bloc_M2471Etiqueteuse".Moteur_Con_En )
      Coil( "Moteur_Con_Entree" )
   END_RUNG
   // the same network as SCL:
   "Moteur_Con_Entree" := "Bloc_M2471Etiqueteuse".Mise_En_Marche AND "Bloc_M2471Etiqueteuse".Moteur_Con_En;
END_REGION

REGION Network 3: moteur Etiquetage
   RUNG wire#powerrail
      Contact( "Bloc_M2471Etiqueteuse".Mise_En_Marche )
      Contact( "Bloc_M2471Etiqueteuse".Moteur_Con_Et )
      Coil( "Moteur_Con_Etiquetage" )
   END_RUNG
   // the same network as SCL:
   "Moteur_Con_Etiquetage" := "Bloc_M2471Etiqueteuse".Mise_En_Marche AND "Bloc_M2471Etiqueteuse".Moteur_Con_Et;
END_REGION

REGION Network 4: Moteur Sortie
   RUNG wire#powerrail
      Contact( "Bloc_M2471Etiqueteuse".Mise_En_Marche )
      Contact( "Bloc_M2471Etiqueteuse".Moteur_Con_So )
      Coil( "Moteur_Con_Sortie" )
   END_RUNG
   // the same network as SCL:
   "Moteur_Con_Sortie" := "Bloc_M2471Etiqueteuse".Mise_En_Marche AND "Bloc_M2471Etiqueteuse".Moteur_Con_So;
END_REGION
END_FUNCTION_BLOCK

FUNCTION_BLOCK "Initialisation"   // FB5, LAD
{ S7_Optimized_Access := 'TRUE' }
VERSION : 0.1
   VAR_TEMP   // added for the SCL form of the ladder/FBD networks
      _w1 : Bool;
      _w2 : Bool;
      _w3 : Bool;
   END_VAR
BEGIN

REGION Network 1 (SCL): Vue Menu et Grand Petit Pot
   IF "Bloc_M2471Etiqueteuse".Vue_Menu = 1 THEN
       "Bloc_M2471Etiqueteuse".Grand_Pot := 0;
       "Bloc_M2471Etiqueteuse".Petit_Pot := 0;
   ELSIF "Bloc_M2471Etiqueteuse".Vue_Grand = 1 THEN
       "Bloc_M2471Etiqueteuse".Grand_Pot := 1;
       "Bloc_M2471Etiqueteuse".Petit_Pot := 0;
   ELSIF "Bloc_M2471Etiqueteuse".Vue_Petit = 1 THEN
       "Bloc_M2471Etiqueteuse".Grand_Pot := 0;
       "Bloc_M2471Etiqueteuse".Petit_Pot := 1;
   END_IF;
END_REGION

REGION Network 2: MCPower
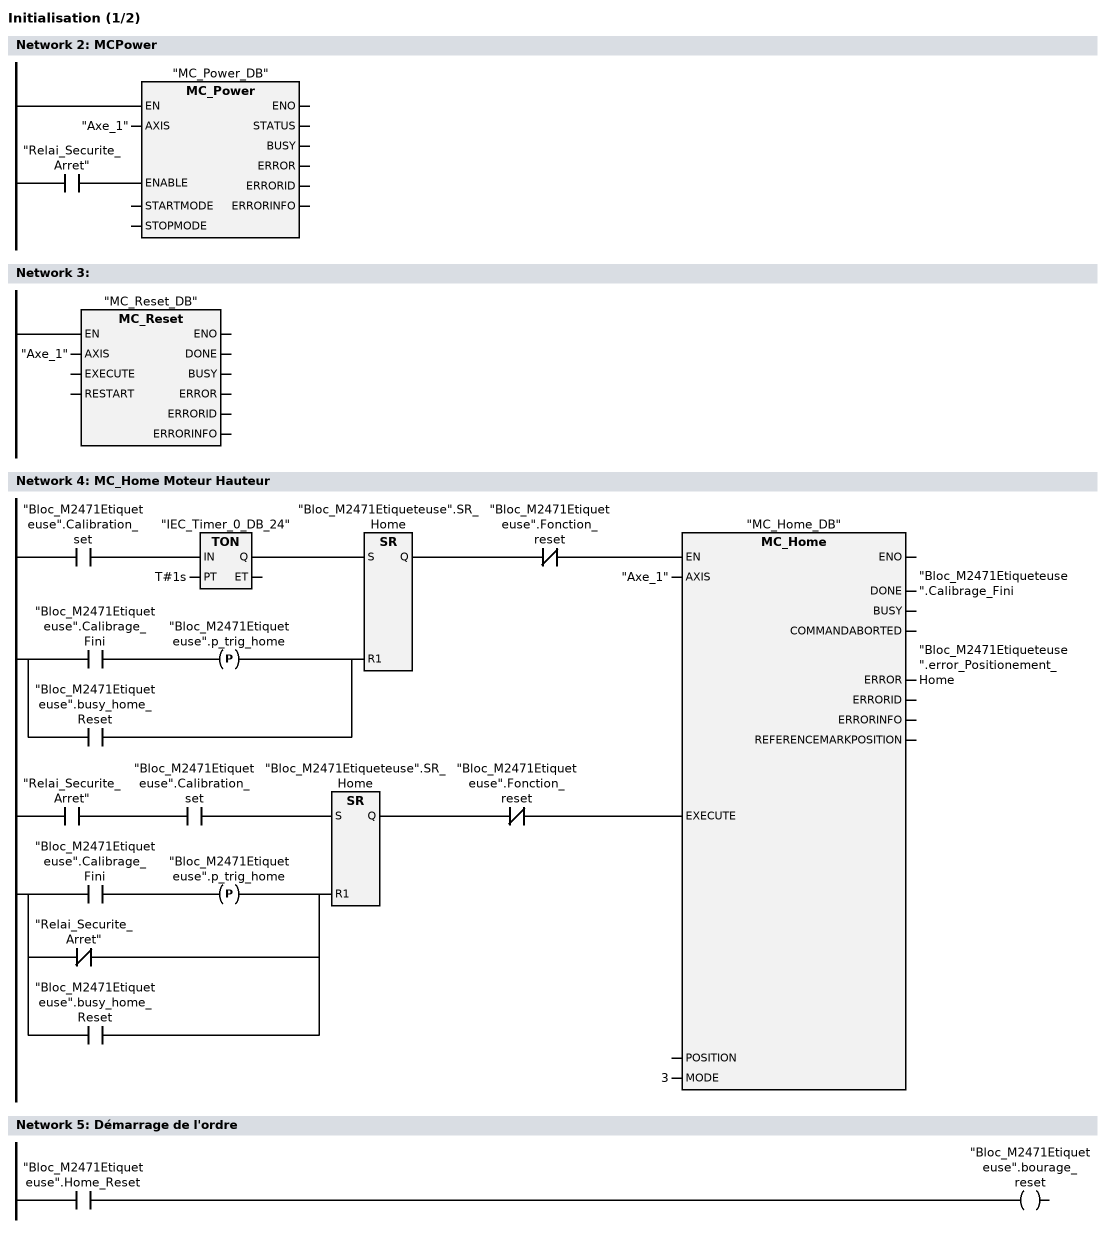
   "MC_Power_DB"(Axis := "Axe_1", Enable := "Relai_Securite_Arret");   // MC_Power
END_REGION

REGION Network 3
   "MC_Reset_DB"(Axis := "Axe_1");   // MC_Reset
END_REGION

REGION Network 4: MC_Home Moteur Hauteur
   "IEC_Timer_0_DB_24".TON(IN := "Bloc_M2471Etiqueteuse".Calibration_set, PT := T#1s);
   #_w1 := "Bloc_M2471Etiqueteuse".Calibrage_Fini AND NOT "Bloc_M2471Etiqueteuse".p_trig_home;   // rising edge
   "Bloc_M2471Etiqueteuse".p_trig_home := "Bloc_M2471Etiqueteuse".Calibrage_Fini;
   IF "IEC_Timer_0_DB_24".Q THEN
       "Bloc_M2471Etiqueteuse".SR_Home := TRUE;   // SR flip-flop
   END_IF;
   IF #_w1 OR "Bloc_M2471Etiqueteuse".busy_home_Reset THEN "Bloc_M2471Etiqueteuse".SR_Home := FALSE; END_IF;
   #_w2 := "Bloc_M2471Etiqueteuse".Calibrage_Fini AND NOT "Bloc_M2471Etiqueteuse".p_trig_home;   // rising edge
   "Bloc_M2471Etiqueteuse".p_trig_home := "Bloc_M2471Etiqueteuse".Calibrage_Fini;
   #_w3 := "Bloc_M2471Etiqueteuse".SR_Home AND NOT "Bloc_M2471Etiqueteuse".Fonction_reset;
   IF "Relai_Securite_Arret" AND "Bloc_M2471Etiqueteuse".Calibration_set THEN
       "Bloc_M2471Etiqueteuse".SR_Home := TRUE;   // SR flip-flop
   END_IF;
   IF #_w2 OR NOT "Relai_Securite_Arret" OR "Bloc_M2471Etiqueteuse".busy_home_Reset THEN
       "Bloc_M2471Etiqueteuse".SR_Home := FALSE;
   END_IF;
   IF #_w3 THEN
       "MC_Home_DB"(Axis := "Axe_1",   // MC_Home
                    Execute := "Bloc_M2471Etiqueteuse".SR_Home AND NOT "Bloc_M2471Etiqueteuse".Fonction_reset,
                    Mode := 3,
                    Done => "Bloc_M2471Etiqueteuse".Calibrage_Fini,
                    Error => "Bloc_M2471Etiqueteuse".error_Positionement_Home);
   END_IF;
END_REGION

REGION Network 5: Démarrage de l'ordre
   RUNG wire#powerrail
      Contact( "Bloc_M2471Etiqueteuse".Home_Reset )
      Coil( "Bloc_M2471Etiqueteuse".bourage_reset )
   END_RUNG
   // the same network as SCL:
   "Bloc_M2471Etiqueteuse".bourage_reset := "Bloc_M2471Etiqueteuse".Home_Reset;
END_REGION

REGION Network 6: Controle Verin Etiquette
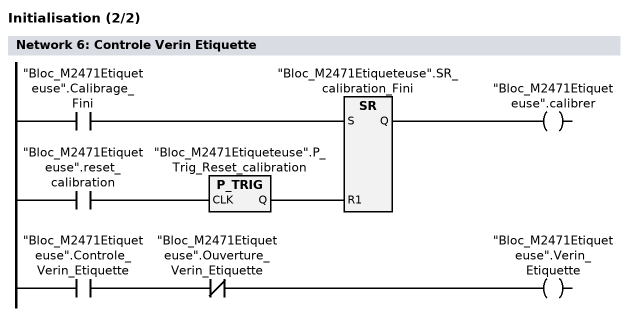
   RUNG wire#powerrail
      Contact( "Bloc_M2471Etiqueteuse".Calibrage_Fini )
      S_SR(operand := "Bloc_M2471Etiqueteuse".SR_calibration_Fini, r1 := wire#w1)
      Coil( "Bloc_M2471Etiqueteuse".calibrer )
   END_RUNG
   RUNG wire#powerrail
      Contact( "Bloc_M2471Etiqueteuse".reset_calibration )
      P_Trig( "Bloc_M2471Etiqueteuse".P_Trig_Reset_calibration )
   END_RUNG wire#w1
   RUNG wire#powerrail
      Contact( "Bloc_M2471Etiqueteuse".Controle_Verin_Etiquette )
      I_Contact( "Bloc_M2471Etiqueteuse".Ouverture_Verin_Etiquette )
      Coil( "Bloc_M2471Etiqueteuse".Verin_Etiquette )
   END_RUNG
   // the same network as SCL:
   #_w1 := "Bloc_M2471Etiqueteuse".reset_calibration AND NOT "Bloc_M2471Etiqueteuse".P_Trig_Reset_calibration;   // rising edge
   "Bloc_M2471Etiqueteuse".P_Trig_Reset_calibration := "Bloc_M2471Etiqueteuse".reset_calibration;
   IF "Bloc_M2471Etiqueteuse".Calibrage_Fini THEN
       "Bloc_M2471Etiqueteuse".SR_calibration_Fini := TRUE;   // SR flip-flop
   END_IF;
   IF #_w1 THEN "Bloc_M2471Etiqueteuse".SR_calibration_Fini := FALSE; END_IF;
   "Bloc_M2471Etiqueteuse".calibrer := "Bloc_M2471Etiqueteuse".SR_calibration_Fini;
   "Bloc_M2471Etiqueteuse".Verin_Etiquette := "Bloc_M2471Etiqueteuse".Controle_Verin_Etiquette AND NOT "Bloc_M2471Etiqueteuse".Ouverture_Verin_Etiquette;
END_REGION

REGION Network 7 (SCL): bouton programe manuel
   IF "Bloc_M2471Etiqueteuse".Bouton_Manuel_5 = 1 THEN
       "Bloc_M2471Etiqueteuse".Valeur_Manuel := 5;
       "Bloc_M2471Etiqueteuse".Bouton_Manuel_10 := 0;
       "Bloc_M2471Etiqueteuse".Bouton_Manuel_25 := 0;

   ELSIF "Bloc_M2471Etiqueteuse".Bouton_Manuel_10 = 1 THEN
       "Bloc_M2471Etiqueteuse".Valeur_Manuel := 10;
       "Bloc_M2471Etiqueteuse".Bouton_Manuel_5 := 0;
       "Bloc_M2471Etiqueteuse".Bouton_Manuel_25 := 0;

   ELSIF "Bloc_M2471Etiqueteuse".Bouton_Manuel_25 = 1 THEN
       "Bloc_M2471Etiqueteuse".Valeur_Manuel := 25;
       "Bloc_M2471Etiqueteuse".Bouton_Manuel_5 := 0;
       "Bloc_M2471Etiqueteuse".Bouton_Manuel_10 := 0;

   END_IF;
END_REGION

REGION Network 8 (SCL): Moteur advance securite coordonne petit et grand >0
   IF "Bloc_M2471Etiqueteuse".Coordone_Grand_Pot > 0 THEN
       "Bloc_M2471Etiqueteuse".valeur_advance_sup_g := 1;
   ELSE
       "Bloc_M2471Etiqueteuse".valeur_advance_sup_g := 0;
   END_IF;
   IF "Bloc_M2471Etiqueteuse".Coordone_Petit_Pot > 0 THEN
       "Bloc_M2471Etiqueteuse".valeur_advance_sup_p := 1;
   ELSE
       "Bloc_M2471Etiqueteuse".valeur_advance_sup_p := 0;
   END_IF;
   IF "Bloc_M2471Etiqueteuse".Vue_Advance =1 AND "Bloc_M2471Etiqueteuse".valeur_advance_sup_g = 1 AND "Bloc_M2471Etiqueteuse".valeur_advance_sup_p = 1 THEN
       "Bloc_M2471Etiqueteuse".Moteur_advance := 1;
   ELSE
       "Bloc_M2471Etiqueteuse".Moteur_advance := 0;
   END_IF;
END_REGION
END_FUNCTION_BLOCK

FUNCTION_BLOCK "Controle_Etiquetage"   // FB6, LAD
{ S7_Optimized_Access := 'TRUE' }
VERSION : 0.1
   VAR_TEMP   // added for the SCL form of the ladder/FBD networks
      _w1 : Bool;
   END_VAR
BEGIN

REGION Network 1 (SCL): Moteur Etiquette On/Off
   IF "Bloc_M2471Etiqueteuse".Etiquetage = true OR "Bloc_M2471Etiqueteuse".Etiquetage_advance OR "Bloc_M2471Etiqueteuse".Etiquetage_comande THEN
       "Bloc_M2471Etiqueteuse".controle_Pwm := TRUE;
   ELSIF "Bloc_M2471Etiqueteuse".Etiquetage_Fini =TRUE OR "Bloc_M2471Etiqueteuse".Vue_Bourage=1  THEN
       "Bloc_M2471Etiqueteuse".controle_Pwm := FALSE;
   END_IF;
END_REGION

REGION Network 2: Capteur Etiquette
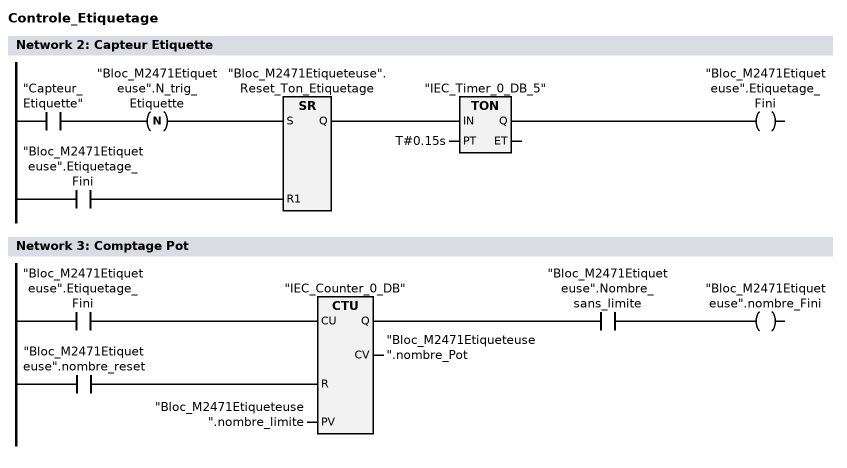
   #_w1 := NOT "Capteur_Etiquette" AND "Bloc_M2471Etiqueteuse".N_trig_Etiquette;   // falling edge
   "Bloc_M2471Etiqueteuse".N_trig_Etiquette := "Capteur_Etiquette";
   IF #_w1 THEN
       "Bloc_M2471Etiqueteuse".Reset_Ton_Etiquetage := TRUE;   // SR flip-flop
   END_IF;
   IF "Bloc_M2471Etiqueteuse".Etiquetage_Fini THEN
       "Bloc_M2471Etiqueteuse".Reset_Ton_Etiquetage := FALSE;
   END_IF;
   "IEC_Timer_0_DB_5".TON(IN := "Bloc_M2471Etiqueteuse".Reset_Ton_Etiquetage, PT := T#0.15s);
   "Bloc_M2471Etiqueteuse".Etiquetage_Fini := "IEC_Timer_0_DB_5".Q;
END_REGION

REGION Network 3: Comptage Pot
   "IEC_Counter_0_DB".CTU(CU := "Bloc_M2471Etiqueteuse".Etiquetage_Fini,
                          R := "Bloc_M2471Etiqueteuse".nombre_reset,
                          PV := "Bloc_M2471Etiqueteuse".nombre_limite,
                          CV => "Bloc_M2471Etiqueteuse".nombre_Pot);
   "Bloc_M2471Etiqueteuse".nombre_Fini := "IEC_Counter_0_DB".Q AND "Bloc_M2471Etiqueteuse".Nombre_sans_limite;
END_REGION
END_FUNCTION_BLOCK

ORGANIZATION_BLOCK "Main_M2471"   // OB1, LAD, ProgramCycle
TITLE = "Main Program Sweep (Cycle)"
{ S7_Optimized_Access := 'TRUE' }
VERSION : 0.1
   VAR_INPUT
      Initial_Call : Bool;   // Initial call of this OB
      Remanence : Bool;   // =True, if remanent data are available
   END_VAR
BEGIN

REGION Network 1: Etat et sécurité
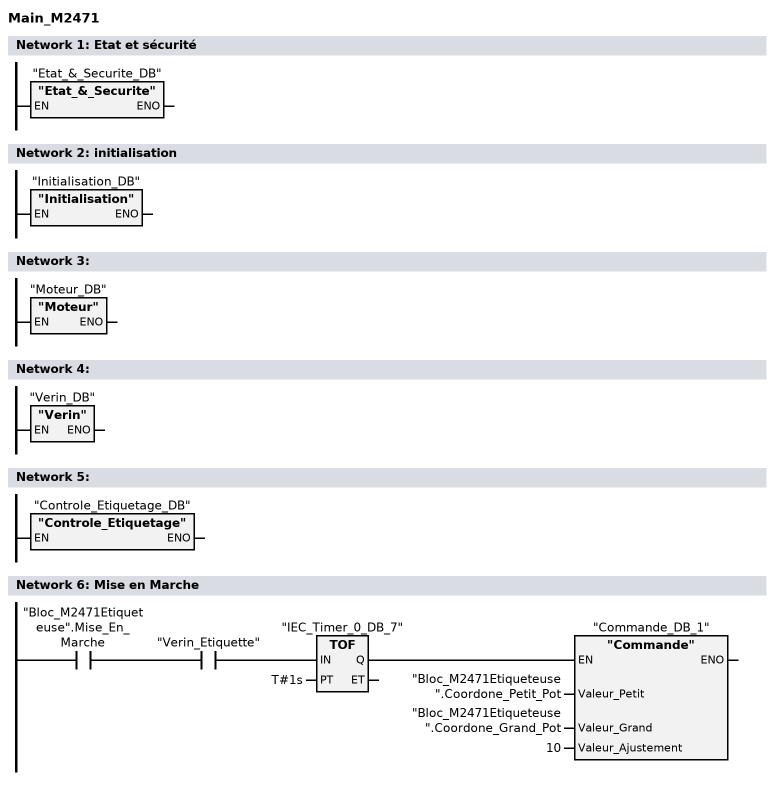
   RUNG wire#powerrail
      "Etat_&_Securite_DB"()
   END_RUNG
   // the same network as SCL:
   "Etat_&_Securite_DB"();   // "Etat_&_Securite"
END_REGION

REGION Network 2: initialisation
   RUNG wire#powerrail
      "Initialisation_DB"()
   END_RUNG
   // the same network as SCL:
   "Initialisation_DB"();   // "Initialisation"
END_REGION

REGION Network 3
   RUNG wire#powerrail
      "Moteur_DB"()
   END_RUNG
   // the same network as SCL:
   "Moteur_DB"();   // "Moteur"
END_REGION

REGION Network 4
   RUNG wire#powerrail
      "Verin_DB"()
   END_RUNG
   // the same network as SCL:
   "Verin_DB"();   // "Verin"
END_REGION

REGION Network 5
   RUNG wire#powerrail
      "Controle_Etiquetage_DB"()
   END_RUNG
   // the same network as SCL:
   "Controle_Etiquetage_DB"();   // "Controle_Etiquetage"
END_REGION

REGION Network 6: Mise en Marche
   "IEC_Timer_0_DB_7".TOF(IN := "Bloc_M2471Etiqueteuse".Mise_En_Marche AND "Verin_Etiquette", PT := T#1s);
   IF "IEC_Timer_0_DB_7".Q THEN
       "Commande_DB_1"(Valeur_Petit := "Bloc_M2471Etiqueteuse".Coordone_Petit_Pot,   // "Commande"
                       Valeur_Grand := "Bloc_M2471Etiqueteuse".Coordone_Grand_Pot,
                       Valeur_Ajustement := 10);
   END_IF;
END_REGION
END_ORGANIZATION_BLOCK

(* ===== HMI "HMI_RT_2" =====
system functions are stored by id; their names below are inferred from use
connection "HMI_Liaison_1": ETHERNET, SMART_S7_1200_OMS

HMI tags "Table de variables standard"
   "Variable_IHM_1" : Int, internal
   "Bloc_M2471Etiqueteuse_Hauteur_Haut" : Bool = PLC Bloc_M2471Etiqueteuse.Hauteur_Haut_Manuel AT %M0.0, 1 s
   "Bloc_M2471Etiqueteuse_Hauteur_Bas" : Bool = PLC Bloc_M2471Etiqueteuse.Hauteur_Bas_Manuel AT %M0.1, 1 s
   "Bloc_M2471Etiqueteuse_Relai_Securite_Etat" : Bool = PLC Bloc_M2471Etiqueteuse.Stop_Etat, 1 s
   "Relai_Securite_Arret" : Bool = PLC Relai_Securite_Arret AT %I0.0, 1 s
   "Bloc_M2471Etiqueteuse_Home" : Bool = PLC Bloc_M2471Etiqueteuse.Calibration_Home, 1 s
   "Bloc_M2471Etiqueteuse_Calibrage_Fini" : Bool = PLC Bloc_M2471Etiqueteuse.Calibrage_Fini, 1 s
   "Bloc_M2471Etiqueteuse_Coordonees_Positionement" : Int = PLC Bloc_M2471Etiqueteuse.Coordonees_Positionement, 1 s
   "Grand_Pot" : Bool = PLC Grand_Pot AT %M1.1, 1 s
   "Bloc_M2471Etiqueteuse_Hauteur_Haut_G_P" : Bool = PLC Bloc_M2471Etiqueteuse.Hauteur_Haut_G_P, 1 s
   "Bloc_M2471Etiqueteuse_Hauteur_Bas_G_P" : Bool = PLC Bloc_M2471Etiqueteuse.Hauteur_Bas_G_P, 1 s
   "Petit_Pot" : Bool = PLC Petit_Pot AT %M1.0, 1 s
   "reset" : Bool = PLC Bloc_M2471Etiqueteuse.Reset AT %I8.6, 1 s
   "retour_Menu" : Bool = PLC retour_Menu AT %M0.5, 1 s
   "Bloc_M2471Etiqueteuse_Reset" : Bool = PLC Bloc_M2471Etiqueteuse.Reset, 1 s
   "Bloc_M2471Etiqueteuse_Grand_Pot" : Bool = PLC Bloc_M2471Etiqueteuse.Grand_Pot, 1 s
   "Bloc_M2471Etiqueteuse_Retour_Menu" : Bool = PLC Bloc_M2471Etiqueteuse.Retour_Menu, 1 s
   "Bloc_M2471Etiqueteuse_Petit_Pot" : Bool = PLC Bloc_M2471Etiqueteuse.Petit_Pot, 1 s
   "Bloc_M2471Etiqueteuse_Calibration" : Bool = PLC Bloc_M2471Etiqueteuse.Calibration_set, 1 s
   "Bloc_M2471Etiqueteuse_Ouverture_Verin_Etiquette" : Bool = PLC Bloc_M2471Etiqueteuse.Ouverture_Verin_Etiquette, 1 s
   "Bloc_M2471Etiqueteuse_Vue_Demarage" : Bool = PLC Bloc_M2471Etiqueteuse.Vue_Demarage, 1 s
   "Bloc_M2471Etiqueteuse_Vue_Menu" : Bool = PLC Bloc_M2471Etiqueteuse.Vue_Menu, 1 s
   "Bloc_M2471Etiqueteuse_Vue_Grand" : Bool = PLC Bloc_M2471Etiqueteuse.Vue_Grand, 1 s
   "Bloc_M2471Etiqueteuse_Vue_Petit" : Bool = PLC Bloc_M2471Etiqueteuse.Vue_Petit, 1 s
   "Bloc_M2471Etiqueteuse_Vue_Manuel" : Bool = PLC Bloc_M2471Etiqueteuse.Vue_Manuel, 1 s
   "Bloc_M2471Etiqueteuse_calibrer" : Bool = PLC Bloc_M2471Etiqueteuse.calibrer, 1 s
   "Bloc_M2471Etiqueteuse_Coordone_Grand_Pot" : Int = PLC Bloc_M2471Etiqueteuse.Coordone_Grand_Pot, 1 s
   "Bloc_M2471Etiqueteuse_Coordone_Petit_Pot" : Int = PLC Bloc_M2471Etiqueteuse.Coordone_Petit_Pot, 1 s
   "Bloc_M2471Etiqueteuse_Coordone_Manuel_Pot" : Int = PLC Bloc_M2471Etiqueteuse.Coordone_Manuel_Pot, 1 s
   "Bloc_M2471Etiqueteuse_N_Trig_Relai" : Bool = PLC Bloc_M2471Etiqueteuse.N_Trig_Relai, 1 s
   "Bloc_M2471Etiqueteuse_Relai_Securite_Etat(1)" : Bool = PLC Bloc_M2471Etiqueteuse.Relai_Securite_Etat, 1 s
   "Bloc_M2471Etiqueteuse_nombre_Pot" : Int = PLC Bloc_M2471Etiqueteuse.nombre_Pot, 1 s
   "Bloc_M2471Etiqueteuse_nombre_limite" : Int = PLC Bloc_M2471Etiqueteuse.nombre_limite, 1 s
   "Bloc_M2471Etiqueteuse_nombre_reset" : Bool = PLC Bloc_M2471Etiqueteuse.nombre_reset, 1 s
   "Bloc_M2471Etiqueteuse_Nombre_sans_limite" : Bool = PLC Bloc_M2471Etiqueteuse.Nombre_sans_limite, 1 s
   "Bloc_M2471Etiqueteuse_Ajustement_Hauteur_G_P" : Bool = PLC Bloc_M2471Etiqueteuse.Ajustement_Hauteur_G_P, 1 s
   "Bloc_M2471Etiqueteuse_Vue_Advance" : Bool = PLC Bloc_M2471Etiqueteuse.Vue_Advance, 1 s
   "Bloc_M2471Etiqueteuse_valeur_Grand_Advance" : Int = PLC Bloc_M2471Etiqueteuse.valeur_Grand_Advance, 1 s
   "Bloc_M2471Etiqueteuse_valeur_advance_sup_p" : Bool = PLC Bloc_M2471Etiqueteuse.valeur_advance_sup_p, 1 s
   "Bloc_M2471Etiqueteuse_valeur_advance_sup_g" : Bool = PLC Bloc_M2471Etiqueteuse.valeur_advance_sup_g, 1 s
   "Bloc_M2471Etiqueteuse_Bouton_Manuel_5" : Bool = PLC Bloc_M2471Etiqueteuse.Bouton_Manuel_5, 1 s
   "Bloc_M2471Etiqueteuse_valeur_Petit_Advance" : Int = PLC Bloc_M2471Etiqueteuse.valeur_Petit_Advance, 1 s
   "Bloc_M2471Etiqueteuse_Confirmation_PP" : Bool = PLC Bloc_M2471Etiqueteuse.Confirmation_PP, 1 s
   "Bloc_M2471Etiqueteuse_Confirmation_GP" : Bool = PLC Bloc_M2471Etiqueteuse.Confirmation_GP, 1 s
   "Bloc_M2471Etiqueteuse_Bouton_Manuel_10" : Bool = PLC Bloc_M2471Etiqueteuse.Bouton_Manuel_10, 1 s
   "Bloc_M2471Etiqueteuse_Bouton_Manuel_25" : Bool = PLC Bloc_M2471Etiqueteuse.Bouton_Manuel_25, 1 s
   "Bloc_M2471Etiqueteuse_Bourage_Done" : Bool = PLC Bloc_M2471Etiqueteuse.Bourage_Done, 1 s
   "Capteur_Verin_Etiquette_Max" : Bool = PLC Capteur_Verin_Etiquette_Max AT %I8.0, 1 s
   "Capteur_Verin_Tete_Min" : Bool = PLC Capteur_Verin_Tete_Min AT %I0.5, 1 s
   "Bloc_M2471Etiqueteuse_validation_securite_1" : Bool = PLC Bloc_M2471Etiqueteuse.validation_securite_1, 1 s
   "Bloc_M2471Etiqueteuse_validation_securite_2" : Bool = PLC Bloc_M2471Etiqueteuse.validation_securite_2, 1 s
   "Bloc_M2471Etiqueteuse_Bourage" : Bool = PLC Bloc_M2471Etiqueteuse.Bourage, 1 s
   "Bloc_M2471Etiqueteuse_Controle_Verin_Etiquette" : Bool = PLC Bloc_M2471Etiqueteuse.Controle_Verin_Etiquette, 1 s
   "Bloc_M2471Etiqueteuse_reset_calibration" : Bool = PLC Bloc_M2471Etiqueteuse.reset_calibration, 1 s
   "Verin_Etiquette" : Bool = PLC Verin_Etiquette AT %Q8.4, 1 s
   "Bloc_M2471Etiqueteuse_Vue_Bourage" : Bool = PLC Bloc_M2471Etiqueteuse.Vue_Bourage, 1 s
   "Bloc_M2471Etiqueteuse_Postionement_reset_error" : Bool = PLC Bloc_M2471Etiqueteuse.Postionement_reset_error, 1 s
   "Bloc_M2471Etiqueteuse_Etiquetage" : Bool = PLC Bloc_M2471Etiqueteuse.Etiquetage, 1 s
   "Bloc_M2471Etiqueteuse_Sortie_1_etiquette" : Bool = PLC Bloc_M2471Etiqueteuse.Sortie_1_etiquette, 1 s
   "Bloc_M2471Etiqueteuse_reset_Manuel_Check" : Bool = PLC Bloc_M2471Etiqueteuse.reset_Manuel_Check, 1 s
   "Bloc_M2471Etiqueteuse_Valeur_manuel_bouton" : Bool = PLC Bloc_M2471Etiqueteuse.Valeur_manuel_bouton, 1 s
   "Bloc_M2471Etiqueteuse_coordoonee_positionement_manuel" : Int = PLC Bloc_M2471Etiqueteuse.coordoonee_positionement_manuel, 1 s
   "Bloc_M2471Etiqueteuse_nouvelle_valeur_manuel" : Int = PLC Bloc_M2471Etiqueteuse.nouvelle_valeur_manuel, 1 s
   "Bloc_M2471Etiqueteuse_comptage_advance_g" : Int = PLC Bloc_M2471Etiqueteuse.comptage_advance_g, 1 s
   "Bloc_M2471Etiqueteuse_comptage_advance_p" : Int = PLC Bloc_M2471Etiqueteuse.comptage_advance_p, 1 s
   "Bloc_M2471Etiqueteuse_reset_count_g" : Bool = PLC Bloc_M2471Etiqueteuse.reset_count_g, 1 s
   "Bloc_M2471Etiqueteuse_reset_count_p" : Bool = PLC Bloc_M2471Etiqueteuse.reset_count_p, 1 s
   "Relai_Secu" : Bool = PLC Relai_Secu AT %Q0.0, 1 s
   "Bloc_M2471Etiqueteuse_error_Positionement" : Bool = PLC Bloc_M2471Etiqueteuse.error_Positionement, 1 s
   "MC_Reset_DB_Execute" : Bool = PLC MC_Reset_DB.Execute, 1 s
   "Bloc_M2471Etiqueteuse_reset_execute" : Bool = PLC Bloc_M2471Etiqueteuse.reset_execute, 1 s

recipe "Hauteur Ø80": Pot Ø80 <- "Bloc_M2471Etiqueteuse_Coordone_Grand_Pot"

recipe "Hateur Ø65": Pot Ø65 <- "Bloc_M2471Etiqueteuse_Coordone_Petit_Pot"

recipe "Hauteur Manuel": Manuel <- "Bloc_M2471Etiqueteuse_coordoonee_positionement_manuel"

Template "Modèle_1" 800x480
   Button "Template_Button" at 714,429 size 71x50; TextOff 'Text'
   Button "Template_Button_1" at 614,429 size 71x50; TextOff 'Text'
   Button "Template_Button_2" at 514,429 size 71x50; TextOff 'Text'
   Button "Template_Button_3" at 414,429 size 71x50; TextOff 'Text'
   Button "Template_Button_4" at 314,429 size 71x50; TextOff 'Text'
   Button "Template_Button_5" at 214,429 size 71x50; TextOff 'Text'
   Button "Template_Button_6" at 114,429 size 71x50; TextOff 'Text'
   Button "Template_Button_7" at 14,429 size 71x50; TextOff 'Text'

screen "02-Menu" 800x480, template "Modèle_1"
   on GenerateScreen: ResetBit("Bloc_M2471Etiqueteuse_Vue_Grand"); ResetBit("Bloc_M2471Etiqueteuse_Vue_Petit"); ResetBit("Bloc_M2471Etiqueteuse_Vue_Manuel"); SetBit("Bloc_M2471Etiqueteuse_Vue_Menu")
   on ClearScreen: ResetBit("Bloc_M2471Etiqueteuse_Vue_Menu")
   GraphicView "Vue de graphique_5" at 0,412 size 798x68; Picture "Graphique_1"
   Button "Bouton_1" at 23,371 size 139x92; TextOff 'Ø80×133mm'
      on Release: ActivateScreen("03-Grand", 0)
      Visibility <- "Verin_Etiquette"
   GraphicView "Vue de graphique_2" at 216,139 size 134x210; Picture "Petit_Pot"
   Button "Bouton_2" at 216,370 size 147x93; TextOff 'Ø65×86mm'
      on Release: ActivateScreen("04-Petit", 0)
      Visibility <- "Verin_Etiquette"
   Button "Bouton_3" at 606,372 size 151x91; TextOff 'Manuel'
      on Release: ActivateScreen("05-Manuel", 0)
      on Press: SetBit("Bloc_M2471Etiqueteuse_Bouton_Manuel_5")
      Visibility <- "Verin_Etiquette"
   GraphicView "Vue de graphique_1" at 21,72 size 173x277; Picture "Grand_Pot_2"
   GraphicView "Vue de graphique_3" at 676,2 size 122x130; Picture "M2471_Logo_Miel_MCT"
   Button "Bouton_4" at 561,22 size 99x88; TextOff 'OFF'
      on Press: ResetBit("Bloc_M2471Etiqueteuse_Relai_Securite_Etat"); ResetBit("Bloc_M2471Etiqueteuse_Ouverture_Verin_Etiquette")
      on Release: ActivateScreen("01-Demarage", 0)
   Button "Bouton_5" at 401,251 size 151x88; TextOff 'Recette'
      on Release: ActivateScreen("07-Recette", 0)
   Button "Bouton_6" at 401,371 size 149x91; TextOff 'Automatique'
      on Release: ActivateScreen("06-Advance", 0)
      Visibility <- "Verin_Etiquette"
   Button "Bouton_7" at 401,134 size 151x101; TextOff 'Vérin Etiquette'
      on Press: InvertBit("Bloc_M2471Etiqueteuse_Ouverture_Verin_Etiquette")
   IOField "Champ d'E/S_4" at 644,153 size 113x50; FormatPattern 999
      ProcessValue <- "Bloc_M2471Etiqueteuse_nombre_Pot"
   TextField "Champ de texte_4" at 615,206 size 142x23; Text 'Etiquetage Total'
   TextField "Champ de texte_1" at 209,37 size 257x35; Text 'M2471 Etiqueteuse'
   TextField "Champ de texte_3" at 108,407 size 356x23; Text 'Veuillez enclencher le Vérin de l'étiquette!'
      Visibility <- "Verin_Etiquette"
   Button "Bouton_8" at 606,250 size 151x89; TextOff 'Sortie 1 Etiquette'
      on Press: SetBit("Bloc_M2471Etiqueteuse_Sortie_1_etiquette")
      on Release: ResetBit("Bloc_M2471Etiqueteuse_Sortie_1_etiquette")
      Visibility <- "Verin_Etiquette"

screen "05-Manuel" 800x480, template "Modèle_1"
   on GenerateScreen: SetBit("Bloc_M2471Etiqueteuse_Vue_Manuel")
   on ClearScreen: ResetBit("Bloc_M2471Etiqueteuse_Vue_Manuel")
   Button "Bouton_3" at 676,146 size 96x83; TextOff 'Retour'
      on Release: ActivateScreen("02-Menu", 0)
   GraphicView "Vue de graphique_1" at 61,47 size 125x168; Picture "Fleche-removebg-preview"
   Button "Bouton_1" at 99,80 size 50x109; TextOff 'Text'
      on Press: SetBit("Bloc_M2471Etiqueteuse_Hauteur_Haut")
      on Release: ResetBit("Bloc_M2471Etiqueteuse_Hauteur_Haut")
   GraphicView "Vue de graphique_2" at 61,227 size 124x169; Picture "Fleche-removebg-preview_1"
   Button "Bouton_2" at 99,254 size 50x107; TextOff 'Text'
      on Press: SetBit("Bloc_M2471Etiqueteuse_Hauteur_Bas")
      on Release: ResetBit("Bloc_M2471Etiqueteuse_Hauteur_Bas")
   GraphicView "Vue de graphique_3" at 676,2 size 122x130; Picture "M2471_Logo_Miel_MCT"
   IOField "Champ d'E/S_1" at 447,57 size 135x53; FormatPattern 999
      on Activate: ResetBit("Bloc_M2471Etiqueteuse_Valeur_manuel_bouton")
      on Deactivate: SetBit("Bloc_M2471Etiqueteuse_Valeur_manuel_bouton")
      ProcessValue <- "Bloc_M2471Etiqueteuse_Coordonees_Positionement"
   Button "Bouton_8" at 384,215 size 57x53; TextOff 'Reset'
      on Release: ResetBit("Bloc_M2471Etiqueteuse_nombre_reset")
      on Press: SetBit("Bloc_M2471Etiqueteuse_nombre_reset")
   TextField "Champ de texte_3" at 364,48 size 76x23; Text 'Hauteur'
   Button "Bouton_4" at 449,205 size 142x68; TextOff 'Comptage Pot'
      on Press: InvertBit("Bloc_M2471Etiqueteuse_Nombre_sans_limite")
      Appearance <- "Bloc_M2471Etiqueteuse_Nombre_sans_limite"
   IOField "Champ d'E/S_4" at 504,292 size 77x32; FormatPattern 999
      ProcessValue <- "Bloc_M2471Etiqueteuse_nombre_Pot"
   IOField "Champ d'E/S_3" at 504,333 size 77x54; FormatPattern 999
      ProcessValue <- "Bloc_M2471Etiqueteuse_nombre_limite"
      Appearance <- "Bloc_M2471Etiqueteuse_Nombre_sans_limite"
   TextField "Champ de texte_1" at 394,348 size 110x23; Text 'Pots Objectif'
   TextField "Champ de texte_2" at 406,297 size 94x23; Text 'Etiquetage'
   Button "Bouton_5" at 234,82 size 83x72; TextOff '+/- 5'
      Appearance <- "Bloc_M2471Etiqueteuse_Bouton_Manuel_5"
      on Press: ResetBit("Bloc_M2471Etiqueteuse_Bouton_Manuel_10"); ResetBit("Bloc_M2471Etiqueteuse_Bouton_Manuel_25")
      on Release: SetBit("Bloc_M2471Etiqueteuse_Bouton_Manuel_5")
   Button "Bouton_6" at 234,174 size 83x72; TextOff '+/- 10'
      Appearance <- "Bloc_M2471Etiqueteuse_Bouton_Manuel_10"
      on Press: ResetBit("Bloc_M2471Etiqueteuse_Bouton_Manuel_5"); ResetBit("Bloc_M2471Etiqueteuse_Bouton_Manuel_25")
      on Release: SetBit("Bloc_M2471Etiqueteuse_Bouton_Manuel_10")
   Button "Bouton_7" at 234,266 size 83x72; TextOff '+/- 25'
      Appearance <- "Bloc_M2471Etiqueteuse_Bouton_Manuel_25"
      on Press: ResetBit("Bloc_M2471Etiqueteuse_Bouton_Manuel_5"); ResetBit("Bloc_M2471Etiqueteuse_Bouton_Manuel_10")
      on Release: SetBit("Bloc_M2471Etiqueteuse_Bouton_Manuel_25")
   TextField "Champ de texte_4" at 364,94 size 75x23; Text 'Max:240'
   TextField "Champ de texte_5" at 364,71 size 50x23; Text 'Min:0'
   GraphicView "Vue de graphique_5" at 0,412 size 798x68; Picture "Graphique_1"
   Button "Bouton_9" at 545,125 size 77x49; TextOff 'set'
      on Release: ResetBit("Bloc_M2471Etiqueteuse_Valeur_manuel_bouton")
      on Press: SetBit("Bloc_M2471Etiqueteuse_Valeur_manuel_bouton")
   IOField "Champ d'E/S_2" at 442,131 size 96x32; FormatPattern 999
      ProcessValue <- "Bloc_M2471Etiqueteuse_nouvelle_valeur_manuel"
   TextField "Champ de texte_6" at 364,137 size 64x23; Text 'Manuel'
   TextField "Champ de texte_7" at 113,95 size 43x23; Text '+'
   TextField "Champ de texte_8" at 117,319 size 43x23; Text '-'

screen "03-Grand" 800x480, template "Modèle_1"
   on GenerateScreen: SetBit("Bloc_M2471Etiqueteuse_Vue_Grand")
   on ClearScreen: ResetBit("Bloc_M2471Etiqueteuse_Vue_Grand")
   GraphicView "Vue de graphique_4" at 28,220 size 124x169; Picture "Fleche-removebg-preview_1"
   GraphicView "Vue de graphique_2" at 28,40 size 125x168; Picture "Fleche-removebg-preview"
   Button "Bouton_3" at 676,157 size 96x70; TextOff 'Retour'
      on Press: SetBit("Bloc_M2471Etiqueteuse_Retour_Menu")
      on Release: ResetBit("Bloc_M2471Etiqueteuse_Retour_Menu"); ActivateScreen("02-Menu", 0)
   GraphicView "Vue de graphique_1" at 210,83 size 190x320; Picture "Grand_Pot_2"
   GraphicView "Vue de graphique_3" at 676,2 size 122x130; Picture "M2471_Logo_Miel_MCT"
   IOField "Champ d'E/S_1" at 532,109 size 84x38; FormatPattern 999
      ProcessValue <- "Bloc_M2471Etiqueteuse_Coordonees_Positionement"
   Button "Bouton_1" at 66,73 size 50x134; TextOff 'Text'
      on Release: ResetBit("Bloc_M2471Etiqueteuse_Hauteur_Haut_G_P")
      on Press: SetBit("Bloc_M2471Etiqueteuse_Hauteur_Haut_G_P")
   Button "Bouton_2" at 66,220 size 50x134; TextOff 'Text'
      on Release: ResetBit("Bloc_M2471Etiqueteuse_Hauteur_Bas_G_P")
      on Press: SetBit("Bloc_M2471Etiqueteuse_Hauteur_Bas_G_P")
   Button "Bouton_8" at 433,184 size 57x53; TextOff 'Reset'
      on Release: ResetBit("Bloc_M2471Etiqueteuse_nombre_reset")
      on Press: SetBit("Bloc_M2471Etiqueteuse_nombre_reset")
   GraphicView "Vue de graphique_5" at 0,412 size 798x68; Picture "Graphique_1"
   TextField "Champ de texte_3" at 439,119 size 76x23; Text 'Hauteur'
   TextField "Champ de texte_4" at 186,31 size 238x23; Text 'POT: Ø86×133mm'
   Button "Bouton_4" at 498,174 size 142x68; TextOff 'Comptage Pot'
      Appearance <- "Bloc_M2471Etiqueteuse_Nombre_sans_limite"
      on Press: InvertBit("Bloc_M2471Etiqueteuse_Nombre_sans_limite")
   IOField "Champ d'E/S_4" at 553,261 size 77x32; FormatPattern 999
      ProcessValue <- "Bloc_M2471Etiqueteuse_nombre_Pot"
   IOField "Champ d'E/S_3" at 553,302 size 77x54; FormatPattern 999
      ProcessValue <- "Bloc_M2471Etiqueteuse_nombre_limite"
      Appearance <- "Bloc_M2471Etiqueteuse_Nombre_sans_limite"
   TextField "Champ de texte_1" at 441,317 size 110x23; Text 'Pots Objectif'
   TextField "Champ de texte_2" at 455,266 size 94x23; Text 'Etiquetage'
   TextField "Champ de texte_5" at 66,96 size 43x23; Text '+10'
   TextField "Champ de texte_6" at 70,312 size 43x23; Text '-10'
   TextField "Champ de texte_7" at 676,226 size 74x23; Text 'MANUEL'

screen "04-Petit" 800x480, template "Modèle_1"
   on GenerateScreen: SetBit("Bloc_M2471Etiqueteuse_Vue_Petit")
   on ClearScreen: ResetBit("Bloc_M2471Etiqueteuse_Vue_Petit")
   GraphicView "Vue de graphique_4" at 37,228 size 124x169; Picture "Fleche-removebg-preview_1"
   GraphicView "Vue de graphique_1" at 37,48 size 125x168; Picture "Fleche-removebg-preview"
   Button "Bouton_3" at 676,154 size 96x101; TextOff 'Retour'
      on Press: SetBit("Bloc_M2471Etiqueteuse_Retour_Menu")
      on Release: ResetBit("Bloc_M2471Etiqueteuse_Retour_Menu"); ActivateScreen("02-Menu", 0)
   GraphicView "Vue de graphique_3" at 676,2 size 122x130; Picture "M2471_Logo_Miel_MCT"
   GraphicView "Vue de graphique_2" at 213,91 size 179x286; Picture "Petit_Pot"
   IOField "Champ d'E/S_1" at 529,102 size 96x32; FormatPattern 999
      ProcessValue <- "Bloc_M2471Etiqueteuse_Coordonees_Positionement"
   Button "Bouton_1" at 75,81 size 50x134; TextOff 'Text'
      on Release: ResetBit("Bloc_M2471Etiqueteuse_Hauteur_Haut_G_P"); ResetBit("Bloc_M2471Etiqueteuse_Ajustement_Hauteur_G_P")
      on Press: SetBit("Bloc_M2471Etiqueteuse_Hauteur_Haut_G_P"); SetBit("Bloc_M2471Etiqueteuse_Ajustement_Hauteur_G_P")
   Button "Bouton_2" at 75,228 size 50x134; TextOff 'Text'
      on Release: ResetBit("Bloc_M2471Etiqueteuse_Hauteur_Bas_G_P"); ResetBit("Bloc_M2471Etiqueteuse_Ajustement_Hauteur_G_P")
      on Press: SetBit("Bloc_M2471Etiqueteuse_Hauteur_Bas_G_P"); SetBit("Bloc_M2471Etiqueteuse_Ajustement_Hauteur_G_P")
   TextField "Champ de texte_1" at 448,111 size 71x23; Text 'Hauteur'
   GraphicView "Vue de graphique_5" at 0,412 size 798x68; Picture "Graphique_1"
   IOField "Champ d'E/S_4" at 553,254 size 77x32; FormatPattern 999
      ProcessValue <- "Bloc_M2471Etiqueteuse_nombre_Pot"
   IOField "Champ d'E/S_3" at 553,295 size 77x54; FormatPattern 999
      ProcessValue <- "Bloc_M2471Etiqueteuse_nombre_limite"
      Appearance <- "Bloc_M2471Etiqueteuse_Nombre_sans_limite"
   TextField "Champ de texte_3" at 441,310 size 110x23; Text 'Pots Objectif'
   TextField "Champ de texte_4" at 455,259 size 94x23; Text 'Etiquetage'
   Button "Bouton_8" at 433,177 size 57x53; TextOff 'Reset'
      on Release: ResetBit("Bloc_M2471Etiqueteuse_nombre_reset")
      on Press: SetBit("Bloc_M2471Etiqueteuse_nombre_reset")
   Button "Bouton_4" at 498,167 size 142x68; TextOff 'Comptage Pot'
      Appearance <- "Bloc_M2471Etiqueteuse_Nombre_sans_limite"
      on Press: InvertBit("Bloc_M2471Etiqueteuse_Nombre_sans_limite")
   TextField "Champ de texte_2" at 197,31 size 228x23; Text 'POT: Ø65×86mm'
   TextField "Champ de texte_5" at 79,103 size 43x23; Text '+10'
   TextField "Champ de texte_6" at 79,313 size 43x23; Text '-10'

screen "01-Demarage" 800x480, template "Modèle_1"
   on GenerateScreen: SetBit("Bloc_M2471Etiqueteuse_Vue_Demarage"); ResetBit("Bloc_M2471Etiqueteuse_Bourage"); ResetBit("Bloc_M2471Etiqueteuse_reset_calibration"); ResetBit("Bloc_M2471Etiqueteuse_Reset"); ResetBit("Bloc_M2471Etiqueteuse_validation_securite_1"); ResetBit("Bloc_M2471Etiqueteuse_validation_securite_2")
   on ClearScreen: ResetBit("Bloc_M2471Etiqueteuse_Vue_Demarage")
   Visibility <- "Bloc_M2471Etiqueteuse_N_Trig_Relai"
   GraphicView "Vue de graphique_5" at 0,412 size 798x68; Picture "Graphique_1"
   GraphicView "Vue de graphique_1" at 413,132 size 203x320; Picture "Grand_Pot_2"
   GraphicView "Vue de graphique_2" at 616,187 size 171x257; Picture "Petit_Pot"
   GraphicView "Vue de graphique_3" at 676,2 size 122x130; Picture "M2471_Logo_Miel_MCT"
   Button "Bouton_1" at 119,177 size 198x147; TextOff 'Start'
      on Press: SetBit("Bloc_M2471Etiqueteuse_Relai_Securite_Etat")
      on Release: ActivateScreen("02-Menu", 0)
      Visibility <- "Bloc_M2471Etiqueteuse_Calibrage_Fini"
   TextField "Champ de texte_1" at 23,23 size 366x48; Text 'M2471_Etiqueteuse'
   TextField "Champ de texte_2" at 23,71 size 43x42; Text 'MPO GRR'
   GraphicView "Vue de graphique_4" at 465,23 size 199x88; Picture "CPNV_Logo"
   TextField "Champ de texte_3" at 112,235 size 223x44; Text 'Appuyez sur le bouton SET Pour Démarrer'
      Visibility <- "Bloc_M2471Etiqueteuse_Relai_Securite_Etat(1)"
   TextField "Champ de texte_4" at 111,286 size 188x23; Text 'Calibration en cours...'
      Visibility <- "Bloc_M2471Etiqueteuse_Calibration"

screen "07-Recette" 800x480
   GraphicView "Vue de graphique_5" at 669,116 size 129x364; Picture "Graphique_1"
   RecipeView "Vue de recette_1" at 0,0 size 677x479
   GraphicView "Vue de graphique_3" at 676,2 size 122x130; Picture "M2471_Logo_Miel_MCT"
   Button "Bouton_3" at 688,186 size 96x107; TextOff 'Retour'
      on Release: ActivateScreen("02-Menu", 0)

screen "06-Advance" 800x480, template "Modèle_1"
   on GenerateScreen: SetBit("Bloc_M2471Etiqueteuse_Vue_Advance")
   on ClearScreen: ResetBit("Bloc_M2471Etiqueteuse_Vue_Advance")
   Button "Bouton_3" at 676,154 size 96x69; TextOff 'Retour'
      on Release: ResetBit("Bloc_M2471Etiqueteuse_Retour_Menu"); ActivateScreen("02-Menu", 0)
      on Press: SetBit("Bloc_M2471Etiqueteuse_Retour_Menu")
   GraphicView "Vue de graphique_3" at 676,2 size 122x130; Picture "M2471_Logo_Miel_MCT"
   GraphicView "Vue de graphique_2" at 239,75 size 169x258; Picture "Petit_Pot"
   TextField "Champ de texte_2" at 676,226 size 111x23; Text 'Automatique'
   IOField "Champ d'E/S_4" at 574,115 size 77x32; FormatPattern 999
      ProcessValue <- "Bloc_M2471Etiqueteuse_nombre_Pot"
   IOField "Champ d'E/S_3" at 574,156 size 77x54; FormatPattern 999
      ProcessValue <- "Bloc_M2471Etiqueteuse_nombre_limite"
      Appearance <- "Bloc_M2471Etiqueteuse_Nombre_sans_limite"
   TextField "Champ de texte_3" at 410,180 size 158x23; Text 'Pots Objectif Total'
   TextField "Champ de texte_4" at 425,118 size 142x23; Text 'Etiquetage Total'
   Button "Bouton_8" at 454,38 size 57x53; TextOff 'Reset'
      on Release: ResetBit("Bloc_M2471Etiqueteuse_nombre_reset")
      on Press: SetBit("Bloc_M2471Etiqueteuse_nombre_reset")
   Button "Bouton_4" at 519,28 size 142x68; TextOff 'Comptage Pot'
      on Press: InvertBit("Bloc_M2471Etiqueteuse_Nombre_sans_limite")
      Appearance <- "Bloc_M2471Etiqueteuse_Nombre_sans_limite"
   GraphicView "Vue de graphique_5" at 2,406 size 798x68; Picture "Graphique_1"
   GraphicView "Vue de graphique_1" at 16,11 size 188x324; Picture "Grand_Pot_2"
   IOField "Champ d'E/S_2" at 270,372 size 99x72; FormatPattern 999
      Appearance <- "Bloc_M2471Etiqueteuse_valeur_advance_sup_p"
      ProcessValue <- "Bloc_M2471Etiqueteuse_Coordone_Petit_Pot"
   TextField "Champ de texte_5" at 233,343 size 171x23; Text 'Hauteur Ø65×86mm'
   TextField "Champ de texte_7" at 26,343 size 181x23; Text 'Hauteur Ø86×133mm'
   IOField "Champ d'E/S_6" at 59,372 size 99x72; FormatPattern 999
      Appearance <- "Bloc_M2471Etiqueteuse_valeur_advance_sup_g"
      ProcessValue <- "Bloc_M2471Etiqueteuse_Coordone_Grand_Pot"
   IOField "Champ d'E/S_1" at 544,333 size 107x48; FormatPattern 999
      ProcessValue <- "Bloc_M2471Etiqueteuse_comptage_advance_g"
   IOField "Champ d'E/S_5" at 544,394 size 107x48; FormatPattern 999
      ProcessValue <- "Bloc_M2471Etiqueteuse_comptage_advance_p"
   TextField "Champ de texte_1" at 413,355 size 131x23; Text 'Etiquetage Ø86'
   TextField "Champ de texte_6" at 412,419 size 131x23; Text 'Etiquetage Ø65'
   Button "Bouton_1" at 665,332 size 115x46; TextOff 'Reset Ø86'
      on Press: SetBit("Bloc_M2471Etiqueteuse_reset_count_g")
      on Release: ResetBit("Bloc_M2471Etiqueteuse_reset_count_g")
   Button "Bouton_2" at 665,394 size 115x47; TextOff 'Reset Ø65'
      on Press: SetBit("Bloc_M2471Etiqueteuse_reset_count_p")
      on Release: ResetBit("Bloc_M2471Etiqueteuse_reset_count_p")

screen "8-Bourage" 800x480, template "Modèle_1"
   Visibility <- "Bloc_M2471Etiqueteuse_N_Trig_Relai"
   on GenerateScreen: ResetBit("Bloc_M2471Etiqueteuse_Calibrage_Fini"); SetBit("Bloc_M2471Etiqueteuse_reset_calibration"); SetBit("Bloc_M2471Etiqueteuse_Reset"); ResetBit("Bloc_M2471Etiqueteuse_Ouverture_Verin_Etiquette"); SetBit("Bloc_M2471Etiqueteuse_Vue_Bourage")
   on ClearScreen: ResetBit("Bloc_M2471Etiqueteuse_Reset"); ResetBit("Bloc_M2471Etiqueteuse_Vue_Bourage")
   GraphicView "Vue de graphique_1" at 465,165 size 151x247; Picture "Grand_Pot_2"
   GraphicView "Vue de graphique_2" at 639,201 size 138x211; Picture "Petit_Pot"
   GraphicView "Vue de graphique_3" at 676,2 size 122x130; Picture "M2471_Logo_Miel_MCT"
   TextField "Champ de texte_1" at 27,23 size 366x48; Text 'M2471_Etiqueteuse'
   TextField "Champ de texte_2" at 27,71 size 43x42; Text 'MPO GRR'
   GraphicView "Vue de graphique_4" at 465,23 size 199x88; Picture "CPNV_Logo"
   GraphicView "Vue de graphique_5" at 0,412 size 798x68; Picture "Graphique_1"
   Button "Bouton_1" at 285,324 size 145x103; TextOff 'Retour'
      Visibility <- "Bloc_M2471Etiqueteuse_Bourage_Done"
      on Release: ActivateScreen("01-Demarage", 0); SetBit("Bloc_M2471Etiqueteuse_Bourage_Done")
      on Press: function_b14e0dd5("MC_Reset_DB_Execute", 0); SetBit("Bloc_M2471Etiqueteuse_reset_execute")
   Circle "Cercle_1" at 29,380 size 48x48
      Appearance <- "Capteur_Verin_Tete_Min"
   Circle "Cercle_2" at 29,303 size 48x48
      Appearance <- "Capteur_Verin_Etiquette_Max"
   Button "Bouton_2" at 29,215 size 75x67; TextOff 'Validé'
      Appearance <- "Bloc_M2471Etiqueteuse_validation_securite_2"
      on Press: InvertBit("Bloc_M2471Etiqueteuse_validation_securite_2")
   Button "Bouton_3" at 29,139 size 75x67; TextOff 'Validé'
      on Press: InvertBit("Bloc_M2471Etiqueteuse_validation_securite_1")
      Appearance <- "Bloc_M2471Etiqueteuse_validation_securite_1"
   TextField "Champ de texte_3" at 105,226 size 200x42; Text 'Aucun Pot dans la zone d'étiquetage'
   TextField "Champ de texte_4" at 108,152 size 208x42; Text 'Système d'étiquetage au dessus du point Home'
   TextField "Champ de texte_5" at 83,328 size 129x23; Text 'Verin Etiquette'
   TextField "Champ de texte_6" at 84,404 size 142x23; Text 'Verin Etiquetage'
*)